                        end = q[:]
                        end[5] += delta
                        if not lower[5] <= end[5] <= upper[5]:
                            alt = q[:]
                            alt[5] -= delta
                            if lower[5] <= alt[5] <= upper[5]:
                                log(f'P{i}：J6 {delta:+d}°超限，改用反方向 {-delta:+d}°（终点位姿不变）。')
                                end, delta = alt, -delta
                            if not lower[5] <= end[5] <= upper[5]:
                                for rewound in _checked_j6_rewinds(q, lower, upper, max_deviation):
                                    if lower[5] <= rewound[5] + delta <= upper[5]:
                                        rewinds.append(rewound[:])
                                        q = rewound
                                        end = q[:]
                                        end[5] += delta
                                        break
                                else:
                                    raise ValueError(f'P{i}：J6 {delta:+d}°超限：反方向与整圈回绕均不可行。')
                        if not _fk_matches(end):
                            raise ValueError(f'P{i}：仅旋转J6无法到达所标注TCP，请检查特异点标记/工具。')
                        # v14d：换向步碰撞时，先试反方向（终点位姿不变），再试整圈回绕——
                        # TCP仿真靠方向枚举能避开这类碰撞，P2P 此前只在超限时才换向。
                        # v14j：反方向终点=当前解−delta（旧代码误算 q−2δ，朝向未翻转、FK 必不匹配，
                        # 15/15 种子全死于此——probe_p14_lookahead.py 坐实）。
                        if _movej_test_cached(q, end, 1) != 0:
                            alt = q[:]
                            alt[5] -= delta
                            flipped = False
                            if lower[5] <= alt[5] <= upper[5] and _fk_matches(alt) and _movej_test_cached(q, alt, 1) == 0:
                                log(f'P{i}：J6 {delta:+d}°扫过障碍，改用反方向 {-delta:+d}°（终点位姿不变）。')
                                end, delta, flipped = alt, -delta, True
                            if not flipped:
                                for rewound in _checked_j6_rewinds(q, lower, upper, max_deviation):
                                    cand = rewound[:]
                                    cand[5] += delta
                                    if lower[5] <= cand[5] <= upper[5] and _fk_matches(cand) and _movej_test_cached(q, cand, 1) == 0:
                                        log(f'P{i}：J6 {delta:+d}°两方向均碰，先整圈回绕再换向。')
                                        rewinds.append(rewound[:])
                                        q, end, flipped = rewound, cand, True
                                        break
                            if not flipped:
                                # v14f：两方向都碰——先切到同位姿的其他 IK 分支（碰撞预检过），
                                # 从那里再换向；途经的构型跳记入 rewinds 由执行层逐跳执行。
                                # v14j：枚举基准改为当前（未翻转）位姿——旧代码误用翻转后 target，
                                # 候选再 ±180 回到未翻转位姿，FK 对 target 永不匹配，结构性必死。
                                for cand in sorted(_ik_branch_candidates(_trajectory_pose(q), q),
                                                   key=lambda c: sum((c[j]-q[j])**2 for j in range(6))):
                                    for sgn in (delta, -delta):
                                        after = cand[:]
                                        after[5] += sgn
                                        if not (lower[5] <= after[5] <= upper[5] and _fk_matches(after)):
                                            continue
                                        if _movej_test_cached(q, cand, 1) == 0 and _movej_test_cached(cand, after, 1) == 0:
                                            log(f'P{i}：J6 ±180°两方向均碰，先切IK分支再换向（rewinds 跳转）。')
                                            rewinds.append(cand[:])
                                            q, end, delta, flipped = cand, after, sgn, True
                                            break
                                    if flipped:
                                        break
                            if not flipped:
                                # v14g：同位姿先 MoveL 到场再换向——MoveL 连续选解给出的构型
                                # 正是 TCP仿真 实测可换向的构型（贪心最近解构型两方向都扫障碍）。
                                lin_end, lin_detail = _linear_path_endpoint(q, target)
                                if lin_end is not None:
                                    pre_waypoints = _linear_waypoints(q, target)
                                    if pre_waypoints:
                                        for sgn in (delta, -delta):
                                            after = lin_end[:]
                                            after[5] += sgn
                                            if not (lower[5] <= after[5] <= upper[5] and _fk_matches(after)):
                                                continue
                                            if _movej_test_cached(lin_end, after, 1) == 0:
                                                log(f'P{i}：J6 两方向均碰，先 MoveL 到场（连续选解构型）再{sgn:+d}°换向。')
                                                plan.append(dict(method='MoveL', joints=lin_end[:], special=False,
                                                                 fallback=False, rewinds=[], j6_delta=None,
                                                                 waypoints=pre_waypoints, p2p_note='换向前MoveL到场'))
                                                q, end, delta, flipped = lin_end[:], after, sgn, True
                                                break
                            if not flipped:
                                raise ValueError(f'P{i}：J6 ±180°换向两方向均碰撞（含回绕/分支/MoveL到场尝试），该构型不可行。')
                        note = ('J6自转%+d°' % delta) if rec.get('spin360', False) else ('J6换向%+d°' % delta)
                    else:
                        target = fanuc_values_to_pose(*rec['values'])
                        # v14h：与前一点同位姿（停顿点，如轨迹7 P7）——不重新选解，
                        # 保持当前构型不动，只往计划里记一个停顿点。
                        if max(abs(_trajectory_pose(q).Pos()[j] - target.Pos()[j]) for j in range(3)) < 1e-3 and \
                           pose_angle(invH(target) * _trajectory_pose(q)) < math.radians(.01):
                            plan.append(dict(method='MoveJ', joints=q[:], special=False, fallback=False,
                                             rewinds=[], j6_delta=None, waypoints=[], p2p_note='同位姿停顿'))
                            continue
                        if not seed_used:
                            end = seed[:]  # v14c：首个TCP点直接采用种子分支（离起点可达性已在种子筛选时验证）
                            seed_used = True
                        else:
                            # v14i：前视——下一个执行点是 ±180 换向时，本点选解必须能完成那次换向
                            #（两方向任一可通行），否则贪心构型会把换向逼成死路。
                            nxt = records[i] if i < len(records) else None
                            lookahead_ok = None
                            if nxt is not None and nxt.get('singular', False) and not nxt.get('spin360', False):
                                nxt_values = nxt['values']
                                def lookahead_ok(cand, _vals=nxt_values, _lower=lower, _upper=upper):
                                    nxt_target = fanuc_values_to_pose(*_vals)
                                    for sgn in (180, -180):
                                        after = cand[:]
                                        after[5] += sgn
                                        if not (_lower[5] <= after[5] <= _upper[5]):
                                            continue
                                        err = invH(nxt_target) * _trajectory_pose(after)
                                        if norm(err.Pos()) > 1e-3 or pose_angle(err) > math.radians(.01):
                                            continue
                                        if _movej_test_cached(cand, after, 1) == 0:
                                            return True
                                    return False
                                log(f'P{i}：前视模式（P{i+1}为±180换向，选解需兼顾换向可行性）。')
                            end = (_nearest_ik_from_current_lookahead(q, target, lookahead_ok)
                                   if lookahead_ok else _nearest_ik_from_current(q, target))
                        note = 'TCP最近解直达'
                        forced_lin = False
                        # v14w24：短直线工作段强制 MoveL——P2→P3 这类 ≤210mm/姿态恒定 的
                        # 贴面平移，工艺不允许 MoveJ 关节弧绕行，直走直线（判据与直发门禁同款）。
                        # 前视夜（下一点±180换向）：直线末端同样具备换向资格才强制，否则回落
                        # MoveJ 前视绑定（保住换向可行性纪律）。
                        _rel = _trajectory_pose(q) * invH(target)
                        _seg_mm_f = norm(_rel.Pos())
                        _force_ok = _seg_mm_f <= MOVL_DIRECT_MAX_MM and pose_angle(_rel) <= math.radians(0.5)
                        # v14w33c：回撤段（TCP y 朝基座 >10mm）且下一点是同位姿换姿 ⇒ 让位 MoveJ
                        # 分支前视（强制 MoveL 的端点分支由直线 IK 连续性锁死，会对下一点无路：
                        # P5→P6→P7 实录 P7 被迫 49 跳细分）。工艺贴面滑移（Δy≈0）不受影响。
                        if _force_ok and i >= 2 and _reorient_next_pose(records, i, rec) is not None:
                            try:
                                _y_prev = float(records[i - 2]['values'][1])
                                if float(rec['values'][1]) - _y_prev > 10.0:
                                    _force_ok = False
                                    log(f'P{i}：回撤段且下一点为同位姿换姿——短直线让位 MoveJ 分支前视（v14w33c）。')
                            except Exception:
                                pass
                        if _force_ok:
                            lin_end_f, lin_detail_f = _linear_path_endpoint(q, target)
                            _lin_ok_f = (lin_end_f is not None
                                         and not _real_interfere_combo(lin_end_f)   # v14w26 组合禁区
                                         and (lookahead_ok is None or lookahead_ok(lin_end_f)))
                            if _lin_ok_f:
                                waypoints = _linear_waypoints(q, target)
                                if waypoints:
                                    end, method, fallback = lin_end_f, 'MoveL', True
                                    note = '短直线强制MoveL'
                                    forced_lin = True
                                    log(f'P{i}：短直线段（{_seg_mm_f:.1f}mm/姿态恒定）按工艺直走 MoveL（不尝试 MoveJ 弧）。')
                            elif lin_end_f is not None:
                                log(f'P{i}：短直线段直线末端无前视换向资格，回落 MoveJ 前视绑定。')
                            else:
                                log(f'P{i}：短直线段 MoveL 不可通行（{lin_detail_f}），回落 MoveJ 尝试。')
                        bound_applied = False
                        # v14j：前视绑定执行——本点是换向前夜：前视选出的构型若弧碰，不得退 MoveL
                        # （连续选解会静默锁回当前族，把死局推迟到换向步才爆——种子13 实证），
                        # 也不得由 v14c 救援收无前视资格的分支；只能换用其他前视合格分支直达，
                        # 全部失败则本构型判死、整段换种子重试。
                        if not forced_lin and lookahead_ok is not None and _movej_test_cached(q, end, 1) != 0:
                            detail_bound = _collision_details()
                            bound = None
                            for cand in sorted(_ik_branch_candidates(target, q),
                                               key=lambda c: sum((c[j]-q[j])**2 for j in range(6))):
                                if lookahead_ok(cand) and _movej_test_cached(q, cand, 1) == 0:
                                    bound = cand
                                    break
                            if bound is not None:
                                end, note, bound_applied = bound[:], '前视绑定避障直达', True
                                log(f'P{i}：前视构型弧碰（{detail_bound}），改用另一前视合格分支直达（前视绑定）。')
                            else:
                                raise ValueError(f'P{i}：MoveJ弧碰撞（{detail_bound}），其余前视合格分支均不可通行；'
                                                 '拒绝退 MoveL（连续选解会丢前视资格），本构型判死。')
                        # v14b：MoveJ 直达弧碰撞时，退回 v13 验证过的 MoveL 直线细分执行。
                        # v14w24：强制 MoveL 段不再尝试/回退 MoveJ（工艺直线优先）。
                        if not forced_lin and not bound_applied and _movej_test_cached(q, end, 1) != 0:
                            detail = _collision_details()
                            lin_end, lin_detail = _linear_path_endpoint(q, target)
                            if lin_end is None:
                                # v14c：直线也碰——枚举该目标全部 IK 分支找可通行 MoveJ（换构型救援）
                                # v14w33b：若下一点是【同位姿纯换姿】，优先选「下一点也能单条 MoveJ 贯通」
                                # 的救援分支（P6→P7 教训：P6 为自避碰选的分支对 P7 无路 ⇒ 49 跳细分拖死执行）。
                                _cands = sorted(_ik_branch_candidates(target, q),
                                                key=lambda c: sum((c[j] - q[j]) ** 2 for j in range(6)))
                                _nxt_pose = None
                                try:
                                    if i < len(records):
                                        _nr = records[i]
                                        if _nr['type'] == 'TCP' and not _nr.get('singular', False):
                                            _va = [float(v) for v in rec['values'][:6]]
                                            _vb = [float(v) for v in _nr['values'][:6]]
                                            if (all(abs(_va[k] - _vb[k]) < 1e-9 for k in range(3))
                                                    and any(abs(_va[k] - _vb[k]) > 1e-9 for k in range(3, 6))):
                                                _nxt_pose = fanuc_values_to_pose(*_nr['values'][:6])
                                except Exception:
                                    _nxt_pose = None
                                rescued = None
                                if _nxt_pose is not None:
                                    for cand in _cands:
                                        if _movej_test_cached(q, cand, 1) != 0:
                                            continue
                                        _ok_nxt = False
                                        for nb in _ik_branch_candidates(_nxt_pose, cand):
                                            if (_real_limit_ok(nb, lower, upper)
                                                    and not _real_interfere_combo(nb)
                                                    and _movej_test_cached(cand, nb, 1) == 0):
                                                _ok_nxt = True
                                                break
                                        if _ok_nxt:
                                            rescued = cand
                                            log(f'P{i}：下一点为同位姿换姿——救援分支带前视，选可与下一点单条 MoveJ 贯通的分支。')
                                            break
                                if rescued is None:
                                    for cand in _cands:
                                        if _movej_test_cached(q, cand, 1) == 0:
                                            rescued = cand
                                            break
                                if rescued is None:
                                    raise ValueError(f'P{i}：MoveJ弧碰撞（{detail}），且MoveL直线也失败：{lin_detail}；'
                                                     '该目标全部IK分支均不可通行。')
                                end, note = rescued[:], 'IK分支救援直达'
                                log(f'P{i}：最近解与直线均碰，切换IK分支救援成功。')
                            else:
                                # v14w33：同位姿/近零长（≤1mm）纯换姿段——MoveL 细分会把 90° 姿态差
                                # 切成数十跳小 MoveJ（10-21 P6→P7 实录 49 跳×每跳断连周期≈3s，
                                # 拖死执行）。优先搜无碰 MoveJ 分支单条直达（分支连续性绑死时
                                # 最近解弧碰≠无解）；搜不到再落回 MoveL 细分兜底。
                                # v14w34：_seg_mm_ro 必须是真实位置差——相对位姿平移模长在原地换姿
                                # 时被旋转杠杆放大（p−R·p，(0,-650,380) 处 90° 即 1064.8mm），
                                # 旧算式使 ≤1mm 门槛从未成立、两个搜索入口从未触发。
                                _pa = _trajectory_pose(q).Pos()
                                _pb = target.Pos()
                                _seg_mm_ro = math.sqrt(sum((_pa[_k] - _pb[_k]) ** 2 for _k in range(3)))
                                reorient_direct = None
                                if _seg_mm_ro <= 1.0:
                                    for cand in sorted(_ik_branch_candidates(target, q),
                                                       key=lambda c: sum((c[j]-q[j])**2 for j in range(6))):
                                        if (not _real_interfere_combo(cand)
                                                and _real_limit_ok(cand, lower, upper)
                                                and (lookahead_ok is None or lookahead_ok(cand))
                                                and _movej_test_cached(q, cand, 1) == 0):
                                            reorient_direct = cand
                                            break
                                if reorient_direct is not None:
                                    end, note = reorient_direct[:], '同位姿换姿MoveJ直达'
                                    method, fallback = 'MoveJ', False
                                    waypoints = []
                                    log(f'P{i}：同位姿换姿——MoveL 细分会碎成数十小段，改用无碰 MoveJ 分支单条直达。')
                                elif _seg_mm_ro <= 1.0 and plan and rec['type'] == 'TCP' and i >= 2:
                                    # v14w33d：回改上一步（已入计划、未执行）为可与本点单条 MoveJ 贯通的
                                    # 分支——上一步若走最近解直达/救援，其分支未必对本点有路（P6→P7 实录）。
                                    # 改关节目标后两跳路径均当场重检，证书完整。
                                    _prev_step = plan[-1]
                                    _prev_q = _prev_step['joints']
                                    _prev_prev = plan[-2]['joints'] if len(plan) >= 2 else saved
                                    _prev_pose = fanuc_values_to_pose(*records[i - 2]['values'][:6])
                                    reorient_direct = None
                                    for c6 in sorted(_ik_branch_candidates(_prev_pose, _prev_prev),
                                                     key=lambda c: sum((c[k] - _prev_q[k]) ** 2 for k in range(6))):
                                        if _real_interfere_combo(c6) or not _real_limit_ok(c6, lower, upper):
                                            continue
                                        if _movej_test_cached(_prev_prev, c6, 1) != 0:
                                            continue
                                        for c7 in sorted(_ik_branch_candidates(target, c6),
                                                         key=lambda c: sum((c[k] - c6[k]) ** 2 for k in range(6))):
                                            if _real_interfere_combo(c7) or not _real_limit_ok(c7, lower, upper):
                                                continue
                                            if lookahead_ok is not None and not lookahead_ok(c7):
                                                continue
                                            if _movej_test_cached(c6, c7, 1) != 0:
                                                continue
                                            _prev_step['joints'] = c6[:]
                                            reorient_direct = c7
                                            break
                                        if reorient_direct is not None:
                                            break
                                    if reorient_direct is not None:
                                        end, note = reorient_direct[:], '同位姿换姿MoveJ直达'
                                        method, fallback = 'MoveJ', False
                                        waypoints = []
                                        log(f'P{i}：回改上一步分支后，本点取得单条 MoveJ 直达（两跳均重检无碰）。')
                                if reorient_direct is not None:
                                    pass   # 已在上方处理
                                else:
                                    waypoints = _linear_waypoints(q, target)
                                    if not waypoints:
                                        raise ValueError(f'P{i}：MoveJ弧碰撞（{detail}），MoveL细分采样失败，拒绝。')
                                    end, method, fallback = lin_end, 'MoveL', True
                                    note = 'MoveJ弧碰退回MoveL细分'
                                    log(f'P{i}：MoveJ弧碰撞（{detail}），改走 MoveL 直线细分（{len(waypoints)} 途经点）。')
                    if not all(lower[j] <= end[j] <= upper[j] for j in range(6)):
                        raise ValueError(f'P{i}：关节超限，J6目标={end[5]:.3f}°。')
                    if method == 'MoveJ' and _movej_test_cached(q, end, 1) != 0:
                        # v14e：普通TCP点最后一级救援——v13 遗产 _obstacle_joint_target
                        # （21候选、肘高排序、限TCP偏离）选避障构型，TCP仿真靠它在同一站过关。
                        try:
                            end = _obstacle_joint_target(q, rec['values'], max_deviation, log)
                            note = '避障选解直达'
                        except ValueError:
                            raise ValueError(f'P{i}：MoveJ路径检查失败（含避障选解）：' + _collision_details())
                        if _movej_test_cached(q, end, 1) != 0:
                            raise ValueError(f'P{i}：MoveJ路径检查失败：' + _collision_details())
                    # v14w25：J6 恰=±360 边界值被控制器 -40006 拒收（10-15 17:26/17:33 实录）。
                    # v14w32：±359.999 内推仍防不住「J6 单轴被丢弃」（10-21 P4 实证：J1~J5 全到、
                    # J6 纹丝停在 180、误差 180°）——改为换 (−180,180] 同角表示（359.999→−0.001），
                    # J6 彻底离开 ±360 邻域。换表示会翻转 MoveJ 弧方向 ⇒ 必须重检路径，不过即报规划错误。
                    # spin360/多圈值（|J6|>360.001）不在此列，防绞坏自转语义。
                    if abs(end[5]) >= 359.999 and abs(end[5]) <= 360.001 and not rec.get('spin360'):
                        _j6n = end[5] - math.copysign(360.0, end[5])
                        log(f'P{i}：J6={end[5]:.3f}° 贴 ±360 边界，换同角表示 {_j6n:.3f}°（v14w32：±359.999 仍被丢轴，彻底离开边界邻域）。')
                        end[5] = _j6n
                        for _wp in waypoints:
                            if abs(_wp[5]) >= 359.999 and abs(_wp[5]) <= 360.001:
                                _wp[5] = _wp[5] - math.copysign(360.0, _wp[5])
                        if method == 'MoveJ' and _movej_test_cached(q, end, 1) != 0:
                            raise ValueError(f'P{i}：J6 换同角表示后 MoveJ 路径碰撞：' + _collision_details())
                    # v14w26：解落入实机自干涉组合区（J4×J5，-40006）——MoveJ 解自动换无碰安全
                    # 分支直达；直线段落区（强制/兜底）整段换种子；无安全分支则判死。
                    if _real_interfere_combo(end):
                        if method == 'MoveJ' and rec['type'] == 'TCP' and not rec.get('singular', False):
                            rescued_if = None
                            for cand_if in sorted(_ik_branch_candidates(target, q),
                                                   key=lambda c: sum((c[j]-q[j])**2 for j in range(6))):
                                if (_real_limit_ok(cand_if, lower, upper)
                                        and not _real_interfere_combo(cand_if)
                                        and _movej_test_cached(q, cand_if, 1) == 0):
                                    rescued_if = cand_if
                                    break
                            if rescued_if is None:
                                raise ValueError(f'P{i}：全部无碰分支均落入实机自干涉组合区'
                                                 f'（|J4|>{REAL_INTERFERE_J4_MAX:.0f} 且 |J5|>{REAL_INTERFERE_J5_MIN:.0f}，-40006 实录区），本构型判死。')
                            log(f'P{i}：预选解落入实机自干涉组合区（J4={end[3]:.1f}°, J5={end[4]:.1f}°），换安全分支直达。')
                            end = rescued_if[:]
                            note = '自干涉安全分支直达'
                        else:
                            raise ValueError(f'P{i}：该步解落入实机自干涉组合区（J4={end[3]:.1f}°, J5={end[4]:.1f}°），换种子重试。')
                    plan.append(dict(method=method, joints=end[:], special=rec.get('singular', False), fallback=False,
                                     rewinds=rewinds, j6_delta=delta,
                                     waypoints=waypoints, p2p_note=note))
                    q = end[:]
                if _continuous_profile_active:
                    previous = saved
                    for number, step in enumerate(plan, 1):
                        if step.get('waypoints'):
                            rel = _trajectory_pose(step['joints']) * invH(_trajectory_pose(previous))
                            if (step['method'] != 'MoveL' or norm(rel.Pos()) > MOVL_DIRECT_MAX_MM
                                    or pose_angle(rel) > math.radians(.5)):
                                raise ValueError(f'P{number}将退回{len(step["waypoints"])}段停走，换入口分支重试。')
                        previous = step['joints']
                log('逐段规划完成，开始整段碰撞复核（1mm/1°采样，请稍候）…')
                _verify_obstacle_plan(saved, plan)
                _certify_continuous_direct(records, saved, plan, log)
                _preferred_seed = (seed_context, seed)
                log(f'P2P+奇异点整段路径预检通过：{len(plan)}点。')
                return plan
            except ValueError as exc:
                last_seed_error = exc
                log(f'种子 {seed_rank}/{len(seeds)} 在此构型失败（{exc}），换下一构型整段重试…')
        if last_seed_error is not None:
            raise last_seed_error
    finally:
        _continuous_profile_active = False
        robot.setJoints(saved)
        RDK.Render(True)

root = tk.Tk()
root.title("RoboDK - 机械臂运动控制（P2P v15.21）")
root.geometry("1200x750")
root.resizable(True, True)

tk.Label(root, text="Dobot CR5 运动控制", font=("Microsoft YaHei", 16, "bold")).pack(pady=10)

notebook = ttk.Notebook(root)
notebook.pack(fill=tk.BOTH, expand=True, padx=10, pady=5)

# ---- 选项卡 1：单点运动 ----
tab_single = ttk.Frame(notebook)
notebook.add(tab_single, text="单点运动")

frame_coord = tk.LabelFrame(tab_single, text="目标 TCP（Fanuc 格式）")
frame_coord.pack(fill=tk.X, padx=10, pady=10)

names = ["X (mm)", "Y (mm)", "Z (mm)", "Rx (deg)", "Ry (deg)", "Rz (deg)"]
defaults = ["0.000", "-241.500", "1047.000", "-90.000", "0.000", "180.000"]
entries_single = []

for i in range(6):
    tk.Label(frame_coord, text=names[i]).grid(row=0, column=i*2, padx=5, pady=10)
    e = tk.Entry(frame_coord, width=12)
    e.insert(0, defaults[i])
    e.grid(row=0, column=i*2+1, padx=5, pady=10)
    entries_single.append(e)

frame_mtype = tk.Frame(tab_single)
frame_mtype.pack(fill=tk.X, padx=10, pady=5)
move_type = tk.StringVar(value="MoveL")
tk.Radiobutton(frame_mtype, text="MoveL (直线)", variable=move_type, value="MoveL").pack(side=tk.LEFT, padx=10)
tk.Radiobutton(frame_mtype, text="MoveJ (关节)", variable=move_type, value="MoveJ").pack(side=tk.LEFT, padx=10)

btn_single_frame = tk.Frame(tab_single)
btn_single_frame.pack(fill=tk.X, padx=10, pady=5)

def _read_current():
    read_current(entries_single)
def _fill_current():
    fill_current(entries_single)
def _check_ik():
    check_ik_single(entries_single)
def _exec_single():
    execute_single(entries_single, move_type.get())

tk.Button(btn_single_frame, text="读取当前 TCP", command=_read_current, width=15).pack(side=tk.LEFT, padx=3)
tk.Button(btn_single_frame, text="当前 TCP -> 输入框", command=_fill_current, width=20).pack(side=tk.LEFT, padx=3)
tk.Button(btn_single_frame, text="检测可达性", command=_check_ik, width=15, bg="#2196F3", fg="white").pack(side=tk.LEFT, padx=3)
tk.Button(btn_single_frame, text="执行运动", command=_exec_single, width=20,
          font=("Microsoft YaHei", 10, "bold"), bg="#4CAF50", fg="white").pack(side=tk.LEFT, padx=3)


# ---- 选项卡 2：目标关节运动（实机） ----
tab_joint = ttk.Frame(notebook)
notebook.add(tab_joint, text="目标关节运动")

frame_joint = tk.LabelFrame(tab_joint, text="目标关节（deg）")
frame_joint.pack(fill=tk.X, padx=10, pady=10)

joint_names = ["J1 (deg)", "J2 (deg)", "J3 (deg)", "J4 (deg)", "J5 (deg)", "J6 (deg)"]
joint_defaults = ["0.000", "0.000", "0.000", "0.000", "0.000", "0.000"]
entries_joint = []

for i in range(6):
    tk.Label(frame_joint, text=joint_names[i]).grid(row=0, column=i*2, padx=5, pady=10)
    e = tk.Entry(frame_joint, width=12)
    e.insert(0, joint_defaults[i])
    e.grid(row=0, column=i*2+1, padx=5, pady=10)
    entries_joint.append(e)

btn_joint_frame = tk.Frame(tab_joint)
btn_joint_frame.pack(fill=tk.X, padx=10, pady=8)

def _read_current_joint_values():
    read_current_joints(entries_joint)

def _fill_current_joints():
    fill_current_joints(entries_joint)

def _exec_joint():
    execute_joint_target(entries_joint)

def _zero_joints():
    clear_joint_target(entries_joint)

tk.Button(btn_joint_frame, text="读取当前关节", command=_read_current_joint_values, width=14).pack(side=tk.LEFT, padx=3)
tk.Button(btn_joint_frame, text="当前关节 -> 输入框", command=_fill_current_joints, width=20).pack(side=tk.LEFT, padx=3)
tk.Button(btn_joint_frame, text="执行指定关节 MoveJ", command=_exec_joint, width=24,
          font=("Microsoft YaHei", 10, "bold"), bg="#FF9800", fg="white").pack(side=tk.LEFT, padx=3)
tk.Button(btn_joint_frame, text="清零", command=_zero_joints, width=10).pack(side=tk.LEFT, padx=3)

tk.Label(tab_joint,
         text="输入 J1~J6 目标角度（deg）；完整关节路径预检通过后才发送实机 MoveJ。",
         fg="#555555").pack(anchor=tk.W, padx=15, pady=5)
tk.Label(tab_joint,
         text="安全提示：首次测试建议只改变一个关节、改变 5~10°，确认方向和角度定义正确后再进行大角度运动。",
         fg="#C62828").pack(anchor=tk.W, padx=15, pady=2)

# ---- 选项卡 3：连续运动 ----
tab_traj = ttk.Frame(notebook)
notebook.add(tab_traj, text="连续运动")

frame_traj_input = tk.LabelFrame(
    tab_traj,
    text="连续运动点输入：每次输入 1 个 TCP 点或 1 组关节角度，点击“检查并加入”"
)
frame_traj_input.pack(fill=tk.X, padx=10, pady=10)

type_frame = tk.Frame(frame_traj_input)
type_frame.pack(fill=tk.X, padx=8, pady=5)

tk.Label(type_frame, text="点类型：").pack(side=tk.LEFT, padx=3)

traj_type = tk.StringVar(value="TCP")
tk.Radiobutton(
    type_frame, text="TCP（X,Y,Z,Rx,Ry,Rz）",
    variable=traj_type, value="TCP"
).pack(side=tk.LEFT, padx=8)

tk.Radiobutton(
    type_frame, text="关节（J1~J6）",
    variable=traj_type, value="JOINT"
).pack(side=tk.LEFT, padx=8)

traj_names_tcp = ["X", "Y", "Z", "Rx", "Ry", "Rz"]
traj_names_joint = ["J1", "J2", "J3", "J4", "J5", "J6"]

traj_entries = []

# ---- 末端特异点设置 ----
singular_var = tk.BooleanVar(value=False)
j6_direction_var = tk.IntVar(value=180)

singular_frame = tk.Frame(frame_traj_input)
singular_frame.pack(fill=tk.X, padx=8, pady=3)

tk.Checkbutton(
    singular_frame,
    text="末端特异点（跳过IK，仅J6转动）",
    variable=singular_var
).pack(side=tk.LEFT, padx=3)

tk.Label(singular_frame, text="J6方向：").pack(side=tk.LEFT, padx=(15, 3))
tk.Radiobutton(singular_frame, text="+180°", variable=j6_direction_var, value=180).pack(side=tk.LEFT, padx=3)
tk.Radiobutton(singular_frame, text="-180°", variable=j6_direction_var, value=-180).pack(side=tk.LEFT, padx=3)
spin_var = tk.BooleanVar(value=False)
tk.Checkbutton(singular_frame, text="J6自转360°（第二类，六维与前点相同）", variable=spin_var).pack(side=tk.LEFT, padx=3)

# 输入框单独放在 grid 子容器中。
# frame_traj_input 本身使用 pack 管理子控件，不能再直接对它的子控件使用 grid。
traj_value_frame = tk.Frame(frame_traj_input)
traj_value_frame.pack(fill=tk.X, padx=8, pady=5)

for i in range(6):
    tk.Label(
        traj_value_frame,
        text=traj_names_tcp[i]
    ).grid(row=0, column=i * 2, padx=3, pady=8)

    e = tk.Entry(traj_value_frame, width=12)
    e.grid(row=0, column=i * 2 + 1, padx=4, pady=8)
    traj_entries.append(e)

# 默认先按 TCP 输入显示
tcp_defaults = ["0.000", "-241.500", "1047.000", "-90.000", "0.000", "180.000"]
for e, val in zip(traj_entries, tcp_defaults):
    e.insert(0, val)


def _update_traj_labels_and_defaults():
    """切换 TCP/关节输入时，更新标签和默认值。"""
    names = traj_names_tcp if traj_type.get() == "TCP" else traj_names_joint
    defaults = (
        tcp_defaults
        if traj_type.get() == "TCP"
        else ["0.000"] * 6
    )

    for i, e in enumerate(traj_entries):
        # grid 上的 Label 位于当前列
        for widget in traj_value_frame.grid_slaves(row=0, column=i * 2):
            widget.configure(text=names[i])

        e.delete(0, tk.END)
        e.insert(0, defaults[i])


tk.Radiobutton(
    type_frame, text="TCP（X,Y,Z,Rx,Ry,Rz）",
    variable=traj_type, value="TCP",
    command=_update_traj_labels_and_defaults
).pack_forget()

# 重新建立带 command 的两个单选按钮
for widget in list(type_frame.pack_slaves()):
    if isinstance(widget, tk.Radiobutton):
        widget.destroy()

tk.Radiobutton(
    type_frame, text="TCP（X,Y,Z,Rx,Ry,Rz）",
    variable=traj_type, value="TCP",
    command=_update_traj_labels_and_defaults
).pack(side=tk.LEFT, padx=8)

tk.Radiobutton(
    type_frame, text="关节（J1~J6）",
    variable=traj_type, value="JOINT",
    command=_update_traj_labels_and_defaults
).pack(side=tk.LEFT, padx=8)

btn_traj_input = tk.Frame(tab_traj)
btn_traj_input.pack(fill=tk.X, padx=10, pady=3)

tk.Button(
    btn_traj_input,
    text="检查并加入当前点",
    command=add_and_check_trajectory_point,
    width=22,
    bg="#2196F3",
    fg="white",
    font=("Microsoft YaHei", 10, "bold")
).pack(side=tk.LEFT, padx=3)

tk.Button(
    btn_traj_input,
    text="读取当前TCP并写入",
    command=read_current_tcp_to_traj,
    width=20
).pack(side=tk.LEFT, padx=3)

tk.Button(
    btn_traj_input,
    text="读取当前关节并写入",
    command=read_current_joints_to_traj,
    width=20
).pack(side=tk.LEFT, padx=3)

tk.Button(
    btn_traj_input,
    text="清空当前输入",
    command=clear_trajectory_input,
    width=16
).pack(side=tk.LEFT, padx=3)

tk.Label(
    tab_traj,
    text="加入点时检查格式并保留关节圈数；执行前再进行整段限位、台子和地面碰撞检查。",
    fg="#555555"
).pack(anchor=tk.W, padx=15, pady=3)

frame_record = tk.LabelFrame(
    tab_traj,
    text="已检查通过的连续运动点（按加入顺序执行，可混合 TCP / 关节点）"
)
frame_record.pack(fill=tk.BOTH, expand=True, padx=10, pady=8)

record_text = tk.Text(frame_record, font=("Consolas", 10), height=10)
record_text.pack(fill=tk.BOTH, expand=True, padx=5, pady=5)

btn_record_frame = tk.Frame(tab_traj)
btn_record_frame.pack(fill=tk.X, padx=10, pady=4)

tk.Button(
    btn_record_frame, text="删除最后一点",
    command=delete_last_record, width=15
).pack(side=tk.LEFT, padx=3)

tk.Button(
    btn_record_frame, text="清空全部点",
    command=clear_records, width=15
).pack(side=tk.LEFT, padx=3)

tk.Button(
    btn_record_frame, text="导入轨迹",
    command=import_trajectory, width=14
).pack(side=tk.LEFT, padx=3)

tk.Button(
    btn_record_frame, text="执行整段连续运动",
    command=execute_recorded_trajectory,
    width=24,
    font=("Microsoft YaHei", 10, "bold"),
    bg="#4CAF50", fg="white"
).pack(side=tk.LEFT, padx=3)

tk.Label(
    tab_traj,
    text="执行前按实机当前关节完成台子/地面预检；仅执行已验证方案。驱动报断连时复核实际到位；未到位或其他异常时中止。",
    fg="#555555"
).pack(anchor=tk.W, padx=15, pady=4)

real_deviation_var = tk.StringVar(value="500.0")
frame_deviation = tk.Frame(root)
frame_deviation.pack(fill=tk.X, padx=10, pady=3)
tk.Label(frame_deviation, text="预检MoveJ兜底最大TCP偏离(mm)：").pack(side=tk.LEFT)
tk.Entry(frame_deviation, textvariable=real_deviation_var, width=10).pack(side=tk.LEFT)
tk.Label(frame_deviation, text="默认500：与TCP仿真/轨迹7~11验证口径一致；实机速度10 mm/s（v14w25 调慢）").pack(side=tk.LEFT, padx=8)

# v14w24：法兰补偿MOVL 默认开启，勾选框移除（工艺定型）。v14l 实机判决驱动 MOVL 无工具
# 补偿（按法兰执行，无补偿直发已拉黑勿回归）；v14p 将错就错把法兰位姿当笛卡尔目标直发，
# 法兰被精确送达→物理尖端走在认证直线上。v14w36/37：位姿由调用方自算 invH(PoseFrame)*SolveFK
# （动画=认证直线，根治关节弧假碰撞冻死），发送窗口配单位变换（校验/数字=法兰空间）。
# 适用：MoveL 细分段≤210mm 且姿态恒定（v14w35 门禁）；规划/预检/几何零改动；失败指纹照旧即停；净化失败自动回落细分。
real_movldirect_var = tk.BooleanVar(value=True)   # 仅保留变量接口（执行入口读取）；无 GUI 控件

# ---- 日志区 ----
frame_log = tk.LabelFrame(root, text="日志")
frame_log.pack(fill=tk.BOTH, expand=True, padx=10, pady=5)

text_log = scrolledtext.ScrolledText(frame_log, font=("Consolas", 10), height=8)
text_log.pack(fill=tk.BOTH, expand=True, padx=5, pady=5)

# ============================================================
# 启动
# ============================================================
log("机器人: " + robot.Name())
log("程序就绪。" + LOG_VERSION + " ｜ 模式：RUNMODE_RUN_ROBOT + robot.Connect() ｜ 文件日志：" + LOG_PATH)
_ensure_canonical_tool()   # v14w17：启动守护（覆盖"加载了带归零工具的存档"场景）
log("单点：输入坐标 -> 检测可达性 -> 执行 MoveL/MoveJ")
log("目标关节：输入 J1~J6 -> 实机 MoveJ（不经过 TCP/Fanuc 转换和 IK）")
log("连续运动（P2P v15.21）：修改点位后仍启用分支搜索、防停走及逐段重新认证；无法认证的直线在发送运动前停止；130mm TCP。")

def _log_pump():
    try:
        while True:
            text_log.insert(tk.END, _log_queue.get_nowait() + NL)
            text_log.see(tk.END)
    except Exception:
        pass
    root.after(100, _log_pump)


_close_requested = False


def _idle_tool_guard():
    if not _real_running and not _tool_window_depth:
        try:
            if _same_tool_pose(robot.PoseTool(), eye(4)):
                _ensure_canonical_tool()
            if _close_requested:
                root.destroy()
                return
        except Exception as exc:
            _file_log('工具空闲守护失败：' + str(exc))
    root.after(1000, _idle_tool_guard)


def _on_close():
    global _close_requested
    if _real_running:
        _close_requested = True
        log('已请求关闭：等待当前任务结束并恢复 TCP 后关闭窗口，继续保留到位监控。')
        return
    _ensure_canonical_tool()
    root.destroy()


root.protocol('WM_DELETE_WINDOW', _on_close)
root.after(100, _log_pump)
root.after(1000, _idle_tool_guard)
_start_heartbeat()
try:
    root.mainloop()
except BaseException:
    import traceback
    _file_log('FATAL mainloop: ' + traceback.format_exc())
    raise

--- program _TCP仿真_路径预检 ---

--- Python program TCP真实运动_P2P版 ---
# -*- coding: utf-8 -*-
"""
RoboDK 实机运动控制（基于 robodk_movej_diag.py 的成功模式）
- 单点：TCP 输入 -> IK 检测 -> MoveL/MoveJ 执行
- 连续轨迹：与TCP仿真同款（姿态退让、J6特异点±180°/自转360°、避障规划+缓存）
2026-10-09：连续运动逻辑对齐 机械臂TCP仿真_副本.py；预检偏离默认 50→500（与验证口径一致）
模式：RUNMODE_RUN_ROBOT + robot.Connect()
"""

from robodk.robolink import *
from robodk.robomath import *
import tkinter as tk
from tkinter import ttk, scrolledtext, filedialog
import time
import math
import json
import itertools

ROBOT_SPEED = 10.0   # v14w25：20→10 mm/s（用户要求调慢；顺带拉长指令间隔，缓解驱动掉线-重连压力）
CANONICAL_TOOL = (0.0, 0.0, 130.0, 0.0, 0.0, 0.0)   # v14w40：规范工具 182→126（2026-10-23 最终实测 法兰→TCP=126；v14w27~39 为 182、v14w14~w26 为 100）；守护用
NL = chr(10)
import queue as _queue_mod
_log_queue = _queue_mod.Queue()  # 后台线程日志经队列回流主线程，GUI 不冻结
LOG_PATH = r'D:\mydata\glm-workplace\sim_scripts\real_gui_log_p2p.txt'  # P2P版独立日志，不覆盖v13黑匣子
LOG_VERSION = 'v15.22-20261104'   # ★ 版本号规则（用户 2026-11-03 要求）：【每次改动都要升版本号】
                               # v15   ：从 v14w42 更名（J4 150→178 / P9 入禁直发 / Tool-User 实验开关 / 删超长横幅）
                               # v15.1 ：最后防线同角归一化修复（段6 J4=198.78 ≡ −161.22 被误判超限）
                               # v15.2 ：新增 |J4|>150 单独硬禁区（治 P5 的 J4=172.88 姿态自干涉）
                               # v15.3 ：打开 MOVL_SEND_TOOL_USER（直发前发 Tool(0)/User(0)，验证能否根治断断续续）
                               # v15.4 ：收口 MoveJ 加重试（治 P8 停下：收口遇断连没走完 ⇒ 关节残差 2.68° 残留）
                               # v15.5 ：直发+收口后再做【关节校正重试】（治 P8 停下：收口走假断连分支 ⇒ 报"已完成"但关节没到位）
                               # v15.6 ：_require_joints 改【带重试的稳定判定】（治 P8 尾通过 → P9 开头又失败：中间还在微动）
                               # v15.7 ：直发后先等【关节真静止】再做验收/收口（治 P8 的 elbow-flip 假通过/假失败）
                               # v15.8 ：★直发落点【自干涉安全网】—— 控制器自行选解可能落进禁区 ⇒ 立刻回认证构型
                               # v15.9 ：P8 也禁直发（治"选解自由"：J1/J6 同步偏 9.77° = 另一组 IK 解）⇒ P8 走细分
                               # v15.10：_require_joints 失败时【主动发 MoveJ 校正】（根治 P8 后不动：断连分支对 MoveJ 只等静止不等到位）
                               # 下次改动 ⇒ v15.23；标题与下方"连续运动"横幅要同步改
# v14w41：独立命名 TCP/法兰工具；恢复原工具链接并核验，失败停止；空闲守护与延后关闭。
# 历史版本记录（场景坐标并非实时状态）：★ v14w40（2026-10-23 18:09）：工具定案 126——最终实测 法兰→TCP=126，CANONICAL_TOOL/守护恢复值/banner 同步 126（历史：v14w27~39=182、v14w14~26=100）；配套场景 磨砂圆柱 y −860→−886、挡板 y 56→30（整体 −26 抵消工具加长的 26mm 深度偏移），轨迹13 采用 z460 统一版（连续轨迹13_t126_z460.json）——tool126+z460+场景−26 组合实测预检 21/21 PASS。⚠️ 实物圆柱/挡板须同步 −26；面贴滚轮旧坐标全部失效需重解；轨迹14/15 需在新配置下复验。v14w39（2026-10-22 14:31）：flange 窗口（单位变换+藏把手）从「仅包 RPC」扩大到【覆盖整个 settle 生命周期】。v14w38 失败教训：假断连让 MoveL 调用秒抛、窗口当场关闭、把手提前恢复，而真实滑行+RoboDK 本地退化动画仍在跑——本地动画在弧 66% 被碰撞检测掐停（模型冻点 J1≈67 四次实录同一位置）、红显常驻，收口 MoveJ 从撞点姿态发出被 RoboDK 拦死。v14w39 三件套：①窗口=包装层全程（发送+断连恢复+到位等待，补发重试每次重开窗）；②守卫补恢复隐藏态门把手（防 GUI 中杀留下隐藏态污染预检）；③直发 settle 返回后 robot.setJoints 钉模型到认证终点（清残余态双保险）。真直线 1mm 检查 0 碰撞、柜子零报警不变。v14w38：窗口藏把手（范围不足判负）。v14w37：位姿传递+单位变换（P8 TargetReachError 修复）。v14w35：门禁 210。v14w34：_seg_mm_ro 真位置差。其余见前版注释与 MEMORY。
# v14w32（2026-10-21 10:58）：J6 贴 ±360 边界的处置从「±359.999 内推」改为「换 (−180,180] 同角表示」（359.999→−0.001）——10-21 P4 实证：内推值仍被控制器丢 J6 单轴（J1~J5 全到、J6 停在 180、误差 180°）；换表示后当场重检 MoveJ 路径（方向翻转风险）；spin360/|J6|>360.001 不处理。其余=v14w30（阈值5°；v14w31 已撤回）。
# v14w30（2026-10-21 09:31）：MovL 直发到位阈 MOVL_ARRIVE_TOL_DEG 2°→5°——10-21 P8 实证：tool=182+z=380 构型下控制器 ~5mm 固有落点误差映射为关节 2.58°（tool=100 时代仅 0.7~0.9°），卡死在旧 ≤2° 阈值外被误判"疑似未执行"；臂实为完成态（零速/模式5/无报警）。护栏不降级：法兰级粗验收(≤8mm/≤1°)+MoveJ 收口仍在其后罩终点；60s 上限与不重发不变。（v14w31 稳定窗+补发×3 已于 10-21 按用户要求撤回。）
# v14w29（2026-10-20 16:42）：站内 圆柱+挡板 统一后移（远离基座）82mm（用户指令：尖端距圆柱面仅 14mm 太近、易自干涉）——圆柱 pose.y −840→−922、挡板 pose.y 76→−6；同时修正 10-15 起过期的场景注释。轨迹13 六点 z−82 补丁后离线预检 21/21 全绿（含本次场景移动复验）。
# v14w28（2026-10-20 16:15）：网格注释同步（纯注释版，逻辑零改动）——把手网格手术 v4：连接件加长、把手组件整体外移，【把手工作点=法兰前 182mm】，stl=tools\handle_rod_182_v2.stl（站内已换、未保存）。工具仍=182mm。
# v14w27（2026-10-20 15:49）：工具坐标 100→182mm（用户实测【物理工具真实长度】；站内 PoseTool 已同步 [0,0,182]）——CANONICAL_TOOL/守护恢复值/直发注释同步，全部 IK 按 182 解算。⚠️ 轨迹13 有 5 点（P8/P9/P10/P12/P13）在 182 下超臂展无逆解，重新示教前禁实机。
# v14w26（2026-10-15 18:15）：实机自干涉组合区（PoseSelfInterference 的 J4×J5 耦合，-40006 实录）——J4=-115.5×J5=173.1 与 J4=-109.4×J5=171.5 双拒；安全实录 J4=-83.2×J5=177.6。修：规划期禁选 |J4|>100 且 |J5|>165 的组合（MoveJ 解落区自动换无碰安全分支；直线段落区回落；无安全分支则整段换种子）。沿用 v14w25：速度10mm/s、J6±360内推（保留作防御）；v14w24：短直线强制MoveL、直发默认开。
# v14w20：受控补发。v14w19：三角离零域。v14w17：工具守护。工具=182.000（v14w27 起）；把手网格=v4 手术（把手组件外移、工作点 z=182，尖端=TCP，把手端抓手 z∈[174,182]；v14w28 起 stl=handle_rod_182_v2）。
# 场景（2026-10-20 实测，v14w29 圆柱/挡板统一后移82 后）：圆柱（轴∥X 滚轮 R150×H50）世界包络 X[−25,25] Y[−1062,−782] Z[330,610]；挡板世界包络 X[−235,215] Y[−1232,−932] Z[150,900]。10-13 版旧场景注释坐标已废（10-15 起站内多次平移未同步注释，v14w29 起以本行为准）。
# 控制器日志实锤（logs/all/log）：
#   11:38:20 拒收 MovL(-0.000000,-615.371000,300.000000,90.000000,0.000000,-0.000000)
#            → [MovL#820] the type of params is wrong: -30001 —— 这才是 P9 直发 60s 零位移的真凶；
#   15:55:51 单步同目标接受 MovL(0.000000,-615.371000,299.999986,89.999995,-0.000003,0.000000)
#            → return 0，1.1s 到位、法兰验收 5.08mm/0.61° 过。两样本差在【边界形态】：
#            x 负零/极小负、rx 恰=+90.000000、rz 负零（触发器三候选未最终定死，净化同时设防）。
# 修法：直发前 _movl_digit_safe_joints 只在零附近边界区对发送关节微扰（单关节 ≤0.05°、末端 ≲0.6mm
#   ≪ 圆柱真裕度 19.9mm）；到位/法兰验收/MoveJ 收口仍全部对【原始认证关节】判定，收口回认证构型。
#   净化失败 ⇒ 本段自动改走细分途经点（安全回落，不比 v14u 更糟）。
# 备份：…_v14v4_20261013-1608.py.bak（另有 1208 站内导出副本）；v14v/v2/v3 回退项见 P2P_LESSONS.md。
# 旧 v14u 备注：v14t 10:38 复跑判读——P9 起步延迟 >6s，「起点静止」与「完成静止」反馈不可区分，位置对目标才是唯一可靠锚点
# v12 黑匣子：原生崩溃时把 Python 调用栈转储到独立文件（被动，不影响逻辑）
# 注意：faulthandler.enable 只接受文件对象，传路径字符串会 AttributeError（v12 首版踩坑，已被 except 吞掉）
CRASH_PATH = r'D:\mydata\glm-workplace\sim_scripts\real_gui_crash.txt'
try:
    import faulthandler as _fh
    _crash_fp = open(CRASH_PATH, 'a', encoding='utf-8')
    _fh.enable(_crash_fp, all_threads=True)
except Exception:
    pass

def _file_log(s):
    try:
        import io as _io, time as _time
        with _io.open(LOG_PATH, 'a', encoding='utf-8') as f:
            f.write(_time.strftime('%m-%d %H:%M:%S') + ' | ' + str(s) + NL)
    except Exception:
        pass


RDK = Robolink()

def fanuc_to_pose(x, y, z, rx, ry, rz):
    return Fanuc_2_Pose([x, y, z, rx, ry, rz])

def pose_to_fanuc(pose):
    return Pose_2_Fanuc(pose)

# ---- 获取机器人 ----
robot = RDK.Item('Dobot CR5', ITEM_TYPE_ROBOT)
if not robot.Valid():
    raise Exception("未找到机器人")

# ---- 全局变量 ----
text_points = None
text_log = None
record_text = None
entries_single = None
entries_joint = None
move_type = None
trajectory_records = []
_connected = False

# ============================================================
# 日志
# ============================================================
# v12 心跳：每5秒覆写一次小文件（时间戳+pid+日志末行），进程死亡时间一目了然
HEARTBEAT_PATH = r'D:\mydata\glm-workplace\sim_scripts\real_gui_heartbeat.txt'

def _start_heartbeat():
    import threading as _t, time as _time, os as _os, io as _io
    def _beat():
        while True:
            try:
                last = ''
                try:
                    with _io.open(LOG_PATH, 'r', encoding='utf-8') as f:
                        _lines = f.read().splitlines()
                        last = _lines[-1] if _lines else ''
                except Exception:
                    pass
                with _io.open(HEARTBEAT_PATH, 'w', encoding='utf-8') as f:
                    f.write('%s | pid=%d | alive\nlast: %s\n' % (
                        _time.strftime('%m-%d %H:%M:%S'), _os.getpid(), last[:150]))
            except Exception:
                pass
            _time.sleep(5.0)
    _t.Thread(target=_beat, daemon=True, name='gui_heartbeat').start()


def log(s):
    _file_log(s)  # 先落盘：即使后续 print 阻塞，磁盘日志也不受影响
    print(s)
    if text_log:
        try:
            _log_queue.put_nowait(str(s))
        except Exception:
            text_log.insert(tk.END, str(s) + NL)

# ============================================================
# 连接（只连一次，复用）
# ============================================================
def ensure_connected():
    global _connected
    try:
        status, msg = robot.ConnectedState()
        if status != ROBOTCOM_READY:
            if status >= 0:
                log('机器人未就绪，取消执行：' + str(msg))
                return False
            robot.Connect()
            # v14o：固定 1.5s 改为就绪探测（0.3s 轮询，最多 3s）：假断连恢复是每跳尾部
            # 停顿税的一部分；探测到就绪即返回，未就绪语义与旧版一致（返回 False）。
            for _ in range(10):
                time.sleep(0.3)
                status, msg = robot.ConnectedState()
                if status == ROBOTCOM_READY:
                    break
        _connected = status == ROBOTCOM_READY
        if not _connected:
            log('机器人连接未就绪：' + str(msg))
            return False
        RDK.setRunMode(RUNMODE_RUN_ROBOT)
        return True
    except Exception as exc:
        _connected = False
        log('连接失败：' + str(exc))
        return False


# ============================================================
# 解析坐标
# ============================================================
def parse_points():
    if not text_points:
        return []
    raw = text_points.get("1.0", tk.END)
    points = []
    for line in raw.strip().split(NL):
        line = line.strip()
        if not line or line.startswith("#"):
            continue
        try:
            vals = [float(v.strip()) for v in line.split(",")]
            if len(vals) >= 6:
                points.append(vals[:6])
        except ValueError:
            pass
    return points

# ============================================================
# 读取当前位置
# ============================================================
def read_current(entries=None):
    try:
        pose = robot.Pose()
        v = pose_to_fanuc(pose)
        log("")
        log("当前 TCP：X=%.3f Y=%.3f Z=%.3f Rx=%.3f Ry=%.3f Rz=%.3f" % tuple(v[:6]))
    except Exception as e:
        log("读取失败：%s" % e)

def fill_current(entries=None):
    try:
        pose = robot.Pose()
        v = pose_to_fanuc(pose)
        if entries:
            for e, val in zip(entries, v):
                e.delete(0, tk.END)
                e.insert(0, "%.3f" % val)
        log("当前 TCP 已填入")
    except Exception as e:
        log("读取失败：%s" % e)

# ============================================================
# IK 检测
# 注意：SolveIK 显式使用当前 Tool + Reference，和 MoveL/MoveJ 保持一致。
# ============================================================
def check_ik_single(entries=None):
    if not entries:
        return
    try:
        values = [float(e.get()) for e in entries]
    except ValueError:
        log("输入无效")
        return

    x, y, z, rx, ry, rz = values
    target = fanuc_to_pose(x, y, z, rx, ry, rz)
    log("")
    log("目标：X=%.3f Y=%.3f Z=%.3f Rx=%.3f Ry=%.3f Rz=%.3f" % (x, y, z, rx, ry, rz))

    try:
        tool_pose = robot.PoseTool()
        frame_pose = robot.PoseFrame()
        joints = robot.SolveIK(target, tool=tool_pose, reference=frame_pose)
        if joints is None:
            log("IK 不可达")
        else:
            q = joints.list()
            if len(q) < 6:
                log("IK 返回关节数量异常：%d，原始数据=%r" % (len(q), q))
                return
            log("IK 可达")
            log("  关节：J1=%.2f J2=%.2f J3=%.2f J4=%.2f J5=%.2f J6=%.2f" % tuple(q[:6]))
    except Exception as e:
        log("检测失败：%s" % e)

def check_all_ik():
    points = parse_points()
    if not points:
        log("没有有效点")
        return

    log("")
    log("========== 检测全部 %d 个点 ==========" % len(points))
    all_ok = True
    for i, p in enumerate(points):
        try:
            target = fanuc_to_pose(*p)
            joints = robot.SolveIK(target, tool=robot.PoseTool(), reference=robot.PoseFrame())
            if joints is None:
                log("  P%d: 不可达" % (i+1))
                all_ok = False
            else:
                q = joints.list()
                if len(q) < 6:
                    raise ValueError("IK 返回关节数量异常: %d, raw=%r" % (len(q), q))
                log("  P%d: 可达  J1=%.1f J2=%.1f J3=%.1f J4=%.1f J5=%.1f J6=%.1f" % (i+1, *q[:6]))
        except Exception as e:
            log("  P%d: 检测失败 %s" % (i+1, e))
            all_ok = False
    if all_ok:
        log("全部 %d 个点可达" % len(points))
    else:
        log("存在不可达点，执行前整段预检将拒绝不通过的方案")

# ============================================================
# 执行单点
# ============================================================
def execute_single(entries=None, mtype="MoveL"):
    try:
        if not entries:
            return
        values = [float(e.get()) for e in entries]
        _execute_checked_real([dict(type='TCP', values=values)], single_method=mtype)
    except (ValueError, TypeError) as exc:
        log('单点输入无效：' + str(exc))


# ============================================================
# 连续运动：选项卡3直接输入 TCP / 关节点，逐点检查后加入轨迹
# ============================================================
trajectory_records = []
record_text = None
traj_entries = None
traj_type = None
singular_var = None
j6_direction_var = None
spin_var = None


def _parse_six_from_entries(entries, label):
    if not entries or len(entries) != 6:
        log("%s输入框异常：需要 6 个值" % label)
        return None
    try:
        vals = [float(e.get().strip()) for e in entries]
    except (ValueError, AttributeError):
        log("%s输入无效：6 个值必须全部为数字" % label)
        return None
    if not all(math.isfinite(v) for v in vals):
        log("%s输入无效：不能包含 NaN 或无穷值" % label)
        return None
    return vals


def _check_tcp_reachable(vals):
    """检查单个 TCP 点 IK 是否可达，返回 (True, target, joints)。"""
    try:
        target = fanuc_to_pose(*vals)
        tool_pose = robot.PoseTool()
        frame_pose = robot.PoseFrame()
        joints = robot.SolveIK(target, tool=tool_pose, reference=frame_pose)

        if joints is None:
            log("TCP IK：不可达")
            return False, None, None

        q = joints.list()
        if len(q) < 6:
            log("TCP IK：返回关节数量异常：%r" % q)
            return False, None, None

        log("TCP IK：可达")
        log("  IK关节：J1=%.2f J2=%.2f J3=%.2f J4=%.2f J5=%.2f J6=%.2f" % tuple(q[:6]))
        return True, target, q[:6]
    except Exception as e:
        log("TCP IK 检查失败：%s: %s" % (type(e).__name__, e))
        return False, None, None


def _check_tcp_segment_continuous(prev_vals, curr_vals, segment_index, samples=20):
    """检查前一个 TCP 点到当前 TCP 点之间的整段插补路径 IK 连续可达性。

    暂不考虑障碍物，只对 TCP 位姿做线性插值，并对每个采样位姿执行 SolveIK。
    起点和终点也包含在采样检查中。
    """
    if prev_vals is None:
        return True

    log("开始检查 P%d -> P%d 的 TCP 连续 IK（%d 个采样点）" %
        (segment_index - 1, segment_index, samples + 1))

    tool_pose = robot.PoseTool()
    frame_pose = robot.PoseFrame()

    for k in range(samples + 1):
        t = float(k) / float(samples)
        vals = [prev_vals[i] + (curr_vals[i] - prev_vals[i]) * t for i in range(6)]
        try:
            pose = fanuc_to_pose(*vals)
            joints = robot.SolveIK(pose, tool=tool_pose, reference=frame_pose)
            if joints is None:
                log("  P%d -> P%d：第 %d/%d 个采样点 IK 不可达，t=%.3f" %
                    (segment_index - 1, segment_index, k + 1, samples + 1, t))
                log("  TCP：X=%.3f Y=%.3f Z=%.3f Rx=%.3f Ry=%.3f Rz=%.3f" % tuple(vals))
                return False
            q = joints.list()
            if len(q) < 6:
                log("  P%d -> P%d：第 %d 个采样点 IK 返回异常：%r" %
                    (segment_index - 1, segment_index, k + 1, q))
                return False
        except Exception as e:
            log("  P%d -> P%d：第 %d 个采样点 IK 检查失败：%s: %s" %
                (segment_index - 1, segment_index, k + 1, type(e).__name__, e))
            return False

    log("P%d -> P%d：连续 IK 检查通过" % (segment_index - 1, segment_index))
    return True


def _check_joint_reachable(q):
    """兼容旧代码：关节点不做可达性/限位检查，输入合法即可加入。"""
    return True


def refresh_record_list():
    if record_text is None:
        return

    record_text.delete("1.0", tk.END)

    for i, rec in enumerate(trajectory_records, 1):
        kind = rec["type"]
        vals = rec["values"]

        if kind == "TCP":
            if rec.get("spin360", False):
                mark = " [J6自转360° %s]" % ("+" if rec.get("j6_delta", 360) >= 0 else "-")
            elif rec.get("singular", False):
                mark = " [J6特异点 %s180°]" % ("+" if rec.get("j6_delta", 180) >= 0 else "-")
            else:
                mark = ""
            record_text.insert(
                tk.END,
                "P%-3d [TCP]%s   X=%9.3f Y=%9.3f Z=%9.3f Rx=%8.3f Ry=%8.3f Rz=%8.3f%s" %
                (i, mark, *vals, NL)
            )
        else:
            record_text.insert(
                tk.END,
                "P%-3d [JNT]   J1=%8.3f J2=%8.3f J3=%8.3f J4=%8.3f J5=%8.3f J6=%8.3f%s" %
                (i, *vals, NL)
            )


def add_and_check_trajectory_point():
    values = _parse_six_from_entries(traj_entries, traj_type.get())
    if values is None:
        return
    kind = traj_type.get()
    is_singular = kind == 'TCP' and bool(singular_var.get())
    spin = is_singular and bool(spin_var.get())
    sign = 1 if int(j6_direction_var.get()) >= 0 else -1
    rec = dict(type=kind, values=values, singular=is_singular, spin360=spin,
               j6_delta=sign * (360 if spin else 180))
    try:
        records = _validated_records(trajectory_records + [rec])
    except ValueError as exc:
        log('点未加入：' + str(exc))
        return
    trajectory_records[:] = records
    refresh_record_list()
    if spin:
        log('P%d [TCP-J6自转360°]：已加入；执行时 J1~J5 不变，J6 %+d°。' % (len(records), sign * 360))
    else:
        log('点已加入；完整避障预检将在执行前进行。关节圈数按输入保留。')



def _write_values_to_traj_entries(values, label):
    if not traj_entries or len(traj_entries) != 6:
        log("连续运动输入框异常：无法写入当前%s" % label)
        return False
    for e, val in zip(traj_entries, values[:6]):
        e.delete(0, tk.END)
        e.insert(0, "%.3f" % float(val))
    log("当前%s已写入选项卡3输入框" % label)
    return True


def read_current_tcp_to_traj():
    """读取当前 RoboDK TCP，并写入选项卡3的 TCP 输入框。"""
    try:
        pose = robot.Pose()
        vals = pose_to_fanuc(pose)
        log("========== 读取当前 TCP -> 选项卡3 ==========")
        log("X=%+.3f Y=%+.3f Z=%+.3f Rx=%+.3f Ry=%+.3f Rz=%+.3f" % tuple(vals))
        if traj_type.get() != "TCP":
            traj_type.set("TCP")
            _update_traj_labels_and_defaults()
        return _write_values_to_traj_entries(vals, "TCP")
    except Exception as e:
        log("读取当前 TCP 失败：%s: %s" % (type(e).__name__, e))
        return False


def read_current_joints_to_traj():
    """读取 RoboDK Robot Item 当前关节，并写入选项卡3的关节输入框。"""
    q = read_current_joints(None)
    if q is None or len(q) < 6:
        return False
    log("========== 读取当前关节 -> 选项卡3 ==========")
    if traj_type.get() != "JOINT":
        traj_type.set("JOINT")
        _update_traj_labels_and_defaults()
    return _write_values_to_traj_entries(q, "关节")


def clear_trajectory_input():
    if not traj_entries:
        return

    for e in traj_entries:
        e.delete(0, tk.END)

    if traj_type.get() == "TCP":
        defaults = ["0.000", "-241.500", "1047.000", "-90.000", "0.000", "180.000"]
    else:
        defaults = ["0.000"] * 6

    for e, val in zip(traj_entries, defaults):
        e.insert(0, val)




def import_trajectory():
    filepath = filedialog.askopenfilename(title='导入轨迹', defaultextension='.json', filetypes=[('JSON轨迹','*.json'),('所有文件','*.*')])
    if not filepath:
        return
    try:
        with open(filepath, encoding='utf-8') as f:
            records = _validated_records(json.load(f))
        trajectory_records[:] = records
        refresh_record_list()
        log(f'已导入{len(records)}点：{filepath}。执行前将从实机当前关节重新预检。')
    except Exception as exc:
        log('轨迹导入失败：' + str(exc))


def delete_last_record():
    if trajectory_records:
        rec = trajectory_records.pop()
        refresh_record_list()
        log("已删除最后一点：P%d [%s]" %
            (len(trajectory_records) + 1, rec["type"]))
    else:
        log("当前没有可删除的连续运动点")


def clear_records():
    trajectory_records.clear()
    refresh_record_list()
    log("连续运动点列表已清空")


def execute_recorded_trajectory():
    log('【点击】执行整段连续运动：当前列表 %d 点（转后台线程执行，窗口保持响应）' % len(trajectory_records))
    import threading
    def _worker():
        try:
            _execute_checked_real(list(trajectory_records))
        except Exception as exc:
            log('【线程异常】%s: %s' % (type(exc).__name__, exc))
    threading.Thread(target=_worker, daemon=True, name='real_exec').start()



# 保留旧函数名，避免其他代码调用失效。
def execute_trajectory():
    execute_recorded_trajectory()


# ============================================================
# 实机关节运动
# ============================================================
def _joint_values_from_entries(entries):
    """从 GUI 读取 J1~J6 目标角度。单位：deg。"""
    if not entries or len(entries) != 6:
        log("目标关节输入框异常：需要 J1~J6 共 6 个")
        return None
    try:
        q = [float(e.get().strip()) for e in entries]
    except (ValueError, AttributeError):
        log("目标关节输入无效：J1~J6 必须全部填写数字")
        return None
    if not all(math.isfinite(v) for v in q):
        log("目标关节输入无效：不能包含 NaN 或无穷值")
        return None
    return q


def read_current_joints(entries=None):
    """读取 RoboDK Robot Item 当前关节值，并可直接填入 J1~J6 输入框。
    注意：这里读取的是 RoboDK 当前 Robot Item 的关节状态，不调用 CR5 控制器 GetAngle。
    """
    try:
        joints = robot.SimulatorJoints()
        q = list(joints) if hasattr(joints, "__iter__") else [joints]
        if len(q) < 6:
            log("读取当前关节失败：SimulatorJoints 返回 %r" % (q,))
            log("请确认 RoboDK 窗口中的机器人已经连接并显示实时关节角度。")
            return None

        q = q[:6]
        log("")
        log("========== RoboDK 当前关节 ==========")
        log("J1=%+.3f°  J2=%+.3f°  J3=%+.3f°" % tuple(q[:3]))
        log("J4=%+.3f°  J5=%+.3f°  J6=%+.3f°" % tuple(q[3:]))

        if entries and len(entries) == 6:
            for e, val in zip(entries, q):
                e.delete(0, tk.END)
                e.insert(0, "%.3f" % val)
            log("当前关节已填入 J1~J6 输入框")

        return q
    except Exception as e:
        log("读取 RoboDK 当前关节失败：%s: %s" % (type(e).__name__, e))
        return None


def fill_current_joints(entries=None):
    """当前 RoboDK 关节 -> 目标关节输入框。"""
    return read_current_joints(entries)


def execute_joint_target(entries=None):
    q = _joint_values_from_entries(entries)
    if q is not None:
        _execute_checked_real([dict(type='JOINT', values=q)])



def clear_joint_target(entries=None):
    if not entries:
        return
    for e in entries:
        e.delete(0, tk.END)
        e.insert(0, "0.000")
    log("目标关节输入已清零")

# ============================================================
# GUI
# ============================================================

# 与TCP仿真一致的预检核心；仅在仿真模式调用。
fanuc_values_to_pose = fanuc_to_pose
pose_to_fanuc_values = pose_to_fanuc
MOVEJ_FALLBACK_MAX_DEVIATION_MM = 50.0
# 预检缓存（与TCP仿真副本同款）：生命周期=单次预检规划，_enable_obstacle_checks 每次进入预检时清空。

_plan_cache = {}
_preferred_seed = None  # Ordering hint only; never reuse a collision certificate.


def _lazy_valid_seeds(seeds, start):
    """Keep the existing valid-seed order, testing only seeds actually needed.

    If none is reachable, preserve the old fallback to the unfiltered list.
    """
    found = False
    for seed in seeds:
        if seed is None or _movej_test_cached(start, seed, 1) == 0:
            found = True
            yield seed
    if not found:
        yield from seeds

def _cache_key_joints(q):
    return tuple(round(float(v), 3) for v in q[:6])

def _cache_key_pose(pose):
    return tuple(tuple(round(float(v), 6) for v in row) for row in pose.rows)

def _movej_test_cached(start, end, minstep_deg):
    """robot.MoveJ_Test 的缓存包装，返回值与直接调用完全一致。
    成功时与原调用一样把仿真关节停在终点；失败路径的规划器只依赖局部
    关节变量（不读取此时的模型关节状态），无需复现失败的副作用。"""
    key = ('movej_test', _cache_key_joints(start), _cache_key_joints(end),
           round(float(minstep_deg), 6))
    if key not in _plan_cache:
        _plan_cache[key] = robot.MoveJ_Test(start, end, minstep_deg=minstep_deg)
    elif _plan_cache[key] == 0:
        robot.setJoints(list(end[:6]))
    return _plan_cache[key]

def _tcp_target_to_flange(target):
    """输入是参考系中的TCP；IK需要机器人基座系中的法兰位姿。"""
    return robot.PoseFrame() * target * invH(robot.PoseTool())

def _flange_target_description(target):
    flange = _tcp_target_to_flange(target)
    return ('换算后的法兰中心（基座系）XYZ=' +
            str(tuple(round(v, 3) for v in flange.Pos())) +
            ' mm，法兰Z轴方向=' + str(tuple(round(v, 6) for v in flange.VZ())))


def _validated_records(data):
    if not isinstance(data, list) or not data:
        raise ValueError('轨迹必须是非空点列表。')
    result = []
    for i, rec in enumerate(data, 1):
        kind = str(rec.get('type', '')).upper()
        if kind == 'JNT':
            kind = 'JOINT'
        values = [float(v) for v in rec.get('values', [])]
        if kind not in ('TCP', 'JOINT') or len(values) != 6 or not all(math.isfinite(v) for v in values):
            raise ValueError(f'P{i}：类型或六维数值无效。')
        special = bool(rec.get('singular', False)) and kind == 'TCP'
        spin = special and bool(rec.get('spin360', False))
        raw_delta = int(rec.get('j6_delta', 360 if spin else 180)) if special else 0
        if special and (not result or result[-1]['type'] != 'TCP' or result[-1]['singular']):
            raise ValueError(f'P{i}：特异点前序或转向无效。')
        if special:
            if spin:
                if raw_delta not in (-360, 360):
                    raise ValueError(f'P{i}：J6自转方向必须为+360或-360。')
                if max(abs(a - b) for a, b in zip(values, result[-1]['values'])) > 1e-3:
                    raise ValueError(f'P{i}：J6自转360°特异点的六维数值必须与前一个TCP点完全相同。')
            elif raw_delta not in (-180, 180):
                raise ValueError(f'P{i}：J6方向必须为+180或-180。')
        delta = (360 if spin else 180) * (1 if raw_delta >= 0 else -1) if special else 0
        result.append(dict(type=kind, values=values, singular=special, spin360=spin, j6_delta=delta))
    return result


def _controller_feedback():
    # Dobot CR V3: 1440-byte real-time feedback; no command is sent on this socket.
    import socket
    import struct
    host, port, *_ = robot.ConnectionParams()
    if int(port) != 29999:
        raise RuntimeError('当前连接不是已验证的Dobot CR反馈协议。')
    previous = None
    with socket.create_connection((host, 30004), timeout=3.0) as connection:
        deadline = time.monotonic() + 3.0
        for _ in range(2):
            packet = bytearray()
            while len(packet) < 1440:
                remaining = deadline - time.monotonic()
                if remaining <= 0:
                    raise RuntimeError('实机反馈读取超时。')
                connection.settimeout(remaining)
                part = connection.recv(1440 - len(packet))
                if not part:
                    raise RuntimeError('实机反馈连接已关闭。')
                packet.extend(part)
            length = struct.unpack_from('<Q', packet, 0)[0]
            marker = struct.unpack_from('<Q', packet, 48)[0]
            stamp = struct.unpack_from('<Q', packet, 32)[0]
            if length != 1440 or marker != 0x123456789ABCDEF:
                raise RuntimeError('实机反馈帧格式不匹配。')
            if previous is not None and stamp <= previous:
                raise RuntimeError('实机反馈时间戳未更新。')
            previous = stamp
        q = list(struct.unpack_from('<6d', packet, 192))   # ★真实关节角（v10定位，示教器交叉证实）；旧版误读432="连接基准+指令累加"的假值
        velocity = list(struct.unpack_from('<6d', packet, 480))
        mode = struct.unpack_from('<Q', packet, 24)[0]
        if not all(math.isfinite(v) for v in q + velocity):
            raise RuntimeError('实机反馈包含无效关节数值。')
        return q, velocity, mode


def _live_joints():
    if RDK.RunMode() != RUNMODE_RUN_ROBOT:
        raise RuntimeError('当前不是实机执行模式。')
    status, msg = robot.ConnectedState()
    if status != ROBOTCOM_READY:
        raise RuntimeError('机器人未就绪或已断连：' + str(msg))
    q, velocity, mode = _controller_feedback()
    # 阈值由 0.1 放宽到 1.0：实测静止时 J4/J3 的速度估计噪声可达 0.31°/s
    # （六轴角度 8 次采样完全相同），0.1 会把"其实已静止"误判为运动中而中止任务。
    if mode != 5 or max(abs(v) for v in velocity) > 1.0:
        raise RuntimeError('实机未处于使能静止状态，模式=%s。' % mode)
    return q


def _require_joints(expected, _tries=3, _allow_fix=False):
    """校验关节与预检一致（容差 0.5°）；失败时【主动发一条 MoveJ 校正】，仍不行才抛错。

    ★★★ v15.10（2026-11-03）：根治"走到 P8 后不动"。
    根因（读码确认）：`_settle_core` 的断连分支写的是
        `_wait_arrival_then_static(expect_target)`
      · 直发段传了 expect_target ⇒ 会等到目标 ✓
      · **MoveJ 段传的是 None** ⇒ 退化为「只等静止」✗
      ⇒ 指令被断连打断、手臂停在中途 ⇒ 只要「静止」就算完成 ✗
      ⇒ 下一段开头的 _require_joints 发现差 9.77° ⇒ 抛错 ⇒ 停 ✗
    （历史证据：10-13 12:12 / 15:49 / 15:55 三次同样失败，当时 P8 走的是纯 MoveJ，与直发无关 ✗）

    修法：不再是"发现不一致就停"，而是【发一条 MoveJ 到认证关节】把手臂拉回去，再校验。
      · 目标就是预检认证过的关节构型 ⇒ 确定可达 ⇒ 重发安全 ✓
      · 只补一次（_allow_fix=False 时不再递归）⇒ 不会无限循环 ✓
      · 拉回后仍不一致 ⇒ 才抛错 ✓（护栏不放松）
    """
    last = None
    actual = None
    for k in range(_tries):
        actual = _live_joints()
        last = max(abs(a - b) for a, b in zip(actual, expected))
        if last <= 0.5:
            return
        if k < _tries - 1:
            log('关节偏差 %.2f° > 0.5°（第 %d/%d 次）⇒ 等 0.5s 重读（可能仍在微动）'
                % (last, k + 1, _tries))
            time.sleep(0.5)
    if _allow_fix:
        log('关节偏差 %.2f°（目标%s，实测%s）⇒ 主动发 MoveJ 校正到认证关节（v15.10）'
            % (last, ['%.2f' % v for v in expected], ['%.2f' % v for v in (actual or [])]))
        try:
            robot.MoveJ(list(expected))
            time.sleep(1.0)
            _require_joints(expected, _tries=3, _allow_fix=False)
            log('✓ 校正 MoveJ 生效：关节已回到认证构型')
            return
        except Exception as _fix_exc:  # noqa: BLE001
            log('⚠️ 校正 MoveJ 未生效：%s: %s' % (type(_fix_exc).__name__, _fix_exc))
    raise RuntimeError('关节反馈与预检状态不一致（偏差 %.2f°，目标%s，实测%s），停止后续命令。'
                       % (last, ['%.2f' % v for v in expected], ['%.2f' % v for v in (actual or [])]))


def _retreat_orientation_records(records):
    """加工点变姿态前退到 y=-750，变姿态后返回 y=-775。"""
    result = []
    previous = None
    for index, record in enumerate(records, 1):
        current = dict(record, values=record['values'][:])
        current['label'] = f'P{index}'
        if previous and previous['type'] == current['type'] == 'TCP':
            old, new = previous['values'], current['values']
            changed = pose_angle(invH(fanuc_values_to_pose(*old)) * fanuc_values_to_pose(*new)) > math.radians(.01)
            old_work, new_work = abs(old[1] + 775) < .001, abs(new[1] + 775) < .001
            if changed and (old_work or new_work):
                anchor = old if old_work else new
                retreat = dict(type='TCP', values=[anchor[0], -750., anchor[2]] + old[3:], singular=False,
                               label=f'P{index}前退让', require_linear=old_work)
                result.append(retreat)
                turn = dict(current, values=retreat['values'][:3] + new[3:], label=f'P{index}退让位换向')
                result.append(turn)
                current['singular'] = False
                current['require_linear'] = new_work
        result.append(current)
        previous = record
    return result


def _prepare_real_plan(records, start, deviation, single_method=None):
    RDK.setRunMode(RUNMODE_SIMULATE)
    try:
        RDK.Command('Trace', 'Off')
        robot.setJoints(start)
        if single_method is None:
            return _plan_continuous_trajectory(records, deviation, log)
        _enable_obstacle_checks()
        if robot.MoveJ_Test(start, start, minstep_deg=1) != 0:
            raise ValueError('起始姿态碰撞：' + _collision_details())
        values = records[0]['values']
        method, fallback = single_method, False
        if method not in ('MoveJ','MoveL'):
            raise ValueError('未知单点运动类型。')
        end = None
        waypoints = []
        if method == 'MoveL':
            end, _ = _linear_path_endpoint(start, fanuc_to_pose(*values))
            if end is not None:
                # v13：单点 MoveL 同样不信任驱动 MOVL（纯J6自转也一样，关节插值=同一路径），
                # 改细分途经点+MoveJ 执行
                waypoints = _linear_waypoints(start, fanuc_to_pose(*values))
                if waypoints:
                    log('单点 MoveL 改细分执行：%d 个途经点（步长≤%.0fmm）。' % (len(waypoints), LINEAR_SUBSTEP_MM))
                    log('单点 MoveL 途经跳（共%d跳）：%s' % (len(waypoints), [[float('%.2f' % v) for v in w] for w in waypoints]))
        if end is None:
            end = _obstacle_joint_target(start, values, deviation if method=='MoveL' else None)
            fallback, method = method=='MoveL', 'MoveJ'
        plan = [dict(method=method,joints=end,special=False,fallback=fallback,rewinds=[],j6_delta=None,waypoints=waypoints)]
        _verify_obstacle_plan(start, plan)
        return plan
    finally:
        robot.setJoints(start)
        RDK.Render(True)
        RDK.setRunMode(RUNMODE_RUN_ROBOT)  # 旧版 L615 有此行：预检后必须切回实机模式，否则 _live_joints 直接拒执行


def _wait_controller_static(max_wait_s=20.0, vel_threshold=0.5, samples=5, interval=0.3):
    """轮询30004反馈直到六轴静止（连续samples次速度<阈值），返回(关节, 是否静止)。

    v14o：断连分支以 samples=3/interval=0.2 调用（短跳≈1s，5×0.3s 静止确认占每跳
    尾部 ~1.5s，是停顿税大头）；默认 5×0.3s 供正常路径；20s 静止上限（真断连护栏）不动。"""
    t0 = time.time()
    quiet = 0
    last = None
    while time.time() - t0 < max_wait_s:
        actual, velocity, _mode = _controller_feedback()
        last = actual
        if max(abs(v) for v in velocity) < vel_threshold:
            quiet += 1
            if quiet >= samples:
                return last, True
        else:
            quiet = 0
        time.sleep(interval)
    return last, False


class ControllerMotionFault(RuntimeError):
    """A controller state that must never trigger a motion resend."""
    pass


def _wait_arrival_then_static(target_joints, max_wait_s=20.0):
    """v14u：目标锚定的到位等待——直发后不再猜「起步了没」，只等「到没到」。

    背景（v14t 10:38 P9 实测）：直发指令起步延迟可 >6s，让位 6s 耗尽判「未执行」
    停止后，指令仍被控制器自行执行到精确目标（善后实测 J2 +10°/J3 +20°，余轴不动，
    宏未重发）——「起点静止」与「完成静止」在反馈上不可区分，位置对目标才是唯一
    可靠锚点（速度判据出局：三场停时 J4 0.06~0.42°/s 均为低于阈值的保持抖动）。
    本函数：距目标关节 ≤MOVL_ARRIVE_TOL_DEG 且速度<0.5°/s → 到位完成（此时已在
    目标，无需再做常规静止确认）；每 5s 一行进度日志（顺带实测真实延迟）；
    上限 MOVL_ARRIVE_WAIT_S 超时报「疑似未执行」停待判读；不重发铁律不变。
    target_joints=None → 退化为 _wait_controller_static()，行为与原先完全一致。"""
    if target_joints is not None:
        t0 = time.time()
        t_note = t0
        while True:
            fb = _controller_feedback()
            if fb[2] not in (5, 7, 8):
                raise ControllerMotionFault(
                    '控制器反馈模式=%s，停止等待且不补发；目标关节=%s，实际关节=%s。请检查示教器报警。'
                    % (fb[2], target_joints, fb[0]))
            err = max(abs(a - b) for a, b in zip(fb[0], target_joints))
            if err <= MOVL_ARRIVE_TOL_DEG and max(abs(v) for v in fb[1]) < 0.5:
                log('MovL 直发到位确认：距目标关节%.2f°（%.1fs），验收继续。'
                    % (err, time.time() - t0))
                return fb[0], True
            if time.time() - t0 >= MOVL_ARRIVE_WAIT_S:
                raise RuntimeError(
                    'MovL 直发%.0fs仍未到位（距目标关节%.2f°），疑似未执行，停止待判读。'
                    % (MOVL_ARRIVE_WAIT_S, err))
            if time.time() - t_note >= 5.0:
                log('MovL 直发等待到位：%.0fs，距目标关节%.2f°，续等（不重发，上限%.0fs）。'
                    % (time.time() - t0, err, MOVL_ARRIVE_WAIT_S))
                t_note = time.time()
            time.sleep(0.5)
    return _wait_controller_static(max_wait_s=max_wait_s)


MOVE_OFFSET_TOL = 0.5   # 闭环补偿后的到位容差（°）


TCP_TOOL_NAME = 'CR5_TCP_130mm'
FLANGE_TOOL_NAME = '_CR5_FLANGE_DIRECT_TEMP'
_tool_window_depth = 0


def _same_tool_pose(a, b):
    return max(abs(a[r, c] - b[r, c]) for r in range(4) for c in range(4)) < 1e-7


def _named_tool(name, pose):
    matches = [it for it in robot.Childs()
               if it.Type() == ITEM_TYPE_TOOL and it.Name() == name]
    if len(matches) > 1:
        raise RuntimeError('重复 TCP 工具条目：' + name)
    if matches:
        tool = matches[0]
        if not _same_tool_pose(tool.PoseTool(), pose):
            raise RuntimeError('TCP 工具定义不符，停止待核对：' + name)
        return tool
    return robot.AddTool(pose, name)


def _restore_tool(pose, linked_tool=None):
    """Restore the original item link when possible, and never swallow failure."""
    for attempt in range(2):
        try:
            robot.setPoseTool(linked_tool if linked_tool is not None and linked_tool.Valid() else pose)
            if not _same_tool_pose(robot.PoseTool(), pose):
                raise RuntimeError('PoseTool 恢复后读回不一致')
            return
        except Exception as exc:
            if attempt == 1:
                raise RuntimeError('工具恢复失败，禁止继续运动：' + str(exc)) from exc


def _single_move_settle(method, target, require_joints=True, expect_target=None, flange_space=False, _retry=0):
    """发指令并确认到位——v14w39 窗口版入口：flange_space 时单位变换+藏把手覆盖
    【整个 settle 生命周期】（发送+断连恢复+到位等待）。旧版只包 RPC 一次调用：假断连
    抛出时窗口即关、把手提前回来，RoboDK 本地退化动画在弧 66% 被碰撞检测掐停→模型冻在
    撞点、红显常驻→收口 MoveJ 被拦死（10-22 四次实录含 v14w38）。"""
    global _tool_window_depth
    if not flange_space or _tool_window_depth:
        # A controlled retry already runs inside the outer tool window.
        # Only the outer owner may restore the original TCP.
        return _settle_core(method, target, require_joints, expect_target, flange_space, _retry)
    _ensure_canonical_tool()
    _win_tp = robot.PoseTool()
    _win_link = robot.getLink(ITEM_TYPE_TOOL)
    _win_handle = RDK.Item('门把手_bs1')
    _win_visible = _win_handle.Visible() if _win_handle.Valid() else None
    _flange_tool = _named_tool(FLANGE_TOOL_NAME, eye(4))
    _tool_window_depth += 1
    try:
        robot.setPoseTool(_flange_tool)
        if not _same_tool_pose(robot.PoseTool(), eye(4)):
            raise RuntimeError('法兰工具切换失败，未发送运动指令')
        if _win_visible is not None:
            _win_handle.setVisible(False)
        result = _settle_core(method, target, require_joints, expect_target, True, _retry)
        # Synchronize measured joints before restoring the tool and visible mesh.
        actual, is_static = _wait_controller_static()
        if not is_static:
            raise RuntimeError('法兰直发后未确认静止，停止后续命令。')
        robot.setJoints(actual)
        return result
    finally:
        try:
            _restore_tool(_win_tp, _win_link)
        finally:
            _tool_window_depth -= 1
            if _win_visible is not None:
                _win_handle.setVisible(_win_visible)


def _settle_core(method, target, require_joints, expect_target, flange_space=False, _retry=0):
    """发一条运动指令并确认到位（v10：反馈字段已校正）。

    v14r：require_joints=False 仅供 MovL 直发调用点使用——断连分支的关节级 0.5°
    校验让位给外层法兰级粗验收（≤8mm/≤1°）+MoveJ 微纠偏收口（v14q 09:57 实机
    教训：MovL 直发必触发假断连，0.95° 固有残差在断连分支内即被拦停，外层验收
    根本没执行到）。其余护栏不变：20s 静止上限、重连失败仍停。

    v14u：断连分支改目标锚定到位等待 _wait_arrival_then_static——上限 60s 每 5s
    进度日志；超时报「疑似未执行」停。不重发铁律不变。

    v14w37：直发=【法兰位姿传递 + flange_space 单位变换窗口】双件套——
    ①传位姿（调用方 invH(PoseFrame)*SolveFK(净化关节) 自算）：MoveL 的动画按位姿空间
    直线走=认证路径，根治旧 MoveL(关节) 的关节弧动画扫进圆柱假碰撞冻死（10-22 两次实录）；
    ②发送 RPC 窗口内 PoseTool 置单位变换：MoveL(位姿) 的可达校验/语义都按 TCP 空间做，
    不切工具则法兰位姿被当 TCP 反推（P8 反推法兰 z=744 爆臂展 ⇒ TargetReachError，
    10-22 11:18 实录）；单位变换下校验空间=法兰空间，数字逐位=金标准（实证 0 偏差）。
    动画窗口内直线途经点 12/12 无碰撞（单位变换工具下实测）。
    v14w38：窗口内追加隐藏把手——驱动断连瞬间 RoboDK 本地退化关节动画（会撞圆柱的
    那条弧）是三次冻结的真凶；藏把手=对假路径的检测放行（实测弧中点/冻结姿态
    显隐 True/False 翻转），真直线 1mm 检查本来就 0 碰撞。

    v14w20：受控补发（一次性）——驱动连接恰死在发送时刻时 SendJointMovJ 会静默
    丢弃不发送（反汇编：CONNECTED=False 直接 return False；2026-10-15 09:51 P25
    实发：断连后臂停在发送前位置、误差127.8°）。补发条件（全部满足才补，且全程
    至多一次）：①失败 ②30004 独立反馈证明【零位移】（仍在发送前关节 ≤0.5°）
    ③ensure_connected() 重连成功。指令已上线/延迟执行/落点异常的场景均不满足
    ②（有位移）不会触发——保留原「不重发」语义。历史上"晚执行"案例（v14t）
    后经控制器日志证实为面板拖动误判，非队列延迟。

    历史结论：驱动一直正确执行绝对关节目标；真实关节角在偏移192。"""
    try:
        _start_q = None
        try:
            _start_q = _controller_feedback()[0]
        except Exception:
            _start_q = None
        getattr(robot, method)(target)   # v14w39：flange 窗口已上移至 _single_move_settle 包装层
    except StoppedError as exc:
        if str(exc).strip() != 'Robot not connected':
            raise
        # v14o 静默重连：假断连是本环境常态（每条 MoveJ 指令结束后都可能误报）；30004
        # 反馈通道独立于驱动连接，静止确认与重连并行进行，压缩跳间停顿税。
        # 护栏不变：未自然收尾（20s 上限）仍停、落点仍 0.5° 校验、重连失败仍停。
        log('驱动报断连——等待收尾与后台重连并行进行…')
        import threading as _st
        reconnected = []
        def _bg_reconnect():
            for _r in range(3):
                if ensure_connected():
                    reconnected.append(True)
                    return
                time.sleep(1.0)
        _rt = _st.Thread(target=_bg_reconnect, daemon=True, name='silent_reconnect')
        _rt.start()
        # v14u：到位等待下沉在断连分支（MovL 直发永远走本分支——v14s 教训）——
        # 目标锚定：距目标≤2°且静止=完成，不猜起步。非 MovL 直发退化为常规静止确认。
        try:
            actual, is_static = _wait_arrival_then_static(expect_target)
        except RuntimeError as _arr_exc:
            if isinstance(_arr_exc, ControllerMotionFault):
                raise
            # v14w20：直发「疑似未执行」——零位移+重连成功 ⇒ 补发一次（指令未上线实证）
            if (_retry < 1 and _start_q is not None
                    and max(abs(a - b) for a, b in zip(_controller_feedback()[0], _start_q)) <= MOVE_OFFSET_TOL
                    and ensure_connected()):
                log('直发疑似未执行且零位移（仍在起点）——判定指令未上线，补发一次（v14w20）。')
                return _single_move_settle(method, target, require_joints, expect_target,
                                           flange_space, _retry=_retry + 1)
            raise
        if not is_static:
            raise RuntimeError('驱动报断连后等待%.0fs仍未静止，停止。' % 20.0) from exc
        if require_joints:
            err = max(abs(a - b) for a, b in zip(actual, target))
            if err > MOVE_OFFSET_TOL:
                # v14w20：MoveJ 类「断连收尾后未到位」——零位移+重连成功 ⇒ 补发一次
                if (_retry < 1 and _start_q is not None
                        and max(abs(a - b) for a, b in zip(actual, _start_q)) <= MOVE_OFFSET_TOL
                        and ensure_connected()):
                    log('断连后零位移（仍在起点）——判定指令未上线，补发一次（v14w20）。')
                    return _single_move_settle(method, target, require_joints, expect_target,
                                               flange_space, _retry=_retry + 1)
                raise RuntimeError('断连收尾后未到位：目标%s，实测%s（误差%.2f°），停止待判读。'
                                   % (['%.2f' % v for v in target], ['%.2f' % v for v in actual], err)) from exc
        _rt.join(timeout=4.0)
        if not reconnected:
            raise RuntimeError('已到位但驱动重连失败，停止后续指令。') from exc
        log('驱动断连但运动已自然完成到位；已重连驱动，继续。')
        return
    actual, is_static = _wait_controller_static()
    if not is_static:
        raise RuntimeError('指令返回后等待静止超时（20s），停止。')
    if require_joints:
        err = max(abs(a - b) for a, b in zip(actual, target))
        if err > MOVE_OFFSET_TOL:
            raise RuntimeError('落点偏差%.2f°：目标%s，实测%s，停止待判读。'
                               % (err, ['%.2f' % v for v in target], ['%.2f' % v for v in actual]))
    return


MOVE_OFFSET_TOL = 0.5   # 到位容差（°）：反馈字段校正后，超过即停止待判读


# v13（方案B）：驱动 MOVL 执行层已判死（3 次实机断连指纹 + .pyc 反汇编直连无收尾），
# 所有 MoveL 执行全部替换为「细分途经点 + MoveJ」。作业面短段（≤ TRANSIT_DIRECT_MAX_MM）
# 用 MoveL 指令的 1mm 逆解采样出 ≤ LINEAR_SUBSTEP_MM 的途经关节序列，MoveJ 逐跳执行；
# 过渡段长段优先 MoveJ 直达（须过 TCP 偏离≤max_deviation 且整弧 MoveJ_Test 碰撞检查），
# 不满足才退回细分。预检层 MoveL_Test@1mm 保留：仍是「这一段能不能走直线」的权威筛选器。
TRANSIT_DIRECT_MAX_MM = 300.0   # 超过此段长的 TCP 段视为自由空间过渡段，尝试 MoveJ 直达
LINEAR_SUBSTEP_MM = 20.0        # 作业面细分步长：v14m(40mm) 实机碰撞实证弦误差可吃掉真裕度（轴线距199.9-半径180≈19.9mm），回 20mm 安全基准（v14k 两度全通过）；途经点弦误差 <0.5mm

MOVL_DIRECT_MAX_MM = 250.0   # v14w35（10-22）：150→210——150 是 v14p 照当时谱系（最长≈120mm）取的设计余量，非事故判死值；210 覆盖 200mm 工艺段一指令（y=-719 线翻转点→x=-100），留 FP 边界余量。路径背书不变（认证直线+整段复核）；更长直线段仍走细分
# ★★★ v14w（2026-10-13 16:08）：【禁直发名单清空 = 恢复 P9 直发】+ 发送位姿数字净化。
#   v14v4 按点号拦 P9 是在 -30001 真凶查明前的临时措施（且拦下分支会落空——随名单清空，
#   该落空分支变为不可达死码，留档不删）。真凶 = 控制器 MovL 参数校验拒收【参数形态】
#   （-0.000000 / +90.000000 / -0.000000，见 LOG_VERSION 处实录），不是几何、不是段长：
#   同目标 15:55:51 单步直发实证 return 0、1.1s 到位。净化失败 ⇒ 本段自动改走细分（安全回落）。
# 想再拦某点：改回 (9,) 即可（注意拦下分支的落空缺陷仍在，见 P2P_LESSONS.md）。
# ★★★ 2026-11-03：改回 (9,) —— 针对【新根因】"movL not set tool or user"（不是 -30001）
#   实录（控制器日志 11-03 10:33:24 / 10:33:30）：
#     [MovL#859] Motion args is legal!            ← 参数合法（所以不是 -30001）
#     [MovL#878] movL not set tool or user!!!     ← ★ 工具/用户坐标系没设置
#     [CallProcess#275] ret = 73/76 ... return = 0,{}  ← 被接受，但按【默认 tool/user】执行
#   ⇒ RoboDK 的 DobotCR 驱动下发 MovL(x,y,z,rx,ry,rz) 时【不带 tool/user】✗
#     ⇒ 控制器用开机默认值 ⇒ 与脚本"法兰补偿（PoseTool=eye）"的语义不一致 ⇒ 落点偏离（P9 差 11.80°）✗
#   ⇒ 保底：P9 不做直发，直接走【细分途经点路径】（今天 P5 就是这样走完的：13 途经点 ✓）
#   ⇒ 根治手段见下方 MOVL_SEND_TOOL_USER（实验性，默认关）
# ★★★ v15.9（2026-11-03）：P8 也加入禁直发 —— 直发的"选解自由"问题对 P8 同样致命。
#   实录（v15.8, 11:56:09~14）：
#     P8 直发 → 等静止 ✓ → 法兰验收通过（5.71mm/0.32° ✓）→ 收口 MoveJ
#     ⇒ 控制器最后停在【另一组 IK 解】：
#        目标 [68.33, 41.30, 10.92, 37.78, -90, 158.33]
#        实测 [78.10, 36.86, 19.48, 33.66, -90, 168.10]
#        差   +9.77, -4.44, +8.56, -4.12,  0,  +9.77
#     ⇒ J1 与 J6 同步 +9.77° ⇒ 【基座-腕部互相补偿】的同一法兰位姿、另一组解 ✗
#   ⇒ 根因：MovL 只给位姿 ⇒ 控制器自行选 IK 分支 ⇒ 关节构型不可控 ✗
#     （v15.5~v15.8 的等待/重试/安全网都改变不了这一点 ✗）
#   ⇒ 细分路径是【逐关节】走的 ⇒ 不存在选解问题 ⇒ 关节精确 ✓（代价：8 跳 ≈24 秒）
MOVL_DIRECT_BLOCK_POINTS = (9, 11)

# ★ 实验性开关（v15.3 已打开做验证）：直发前先给【控制器】发 Tool(0)/User(0)，
#   让 MovL 明确用 基座系+零工具(法兰)。背景：[MovL#878] movL not set tool or user!!!
#   ⇒ 控制器没收到 tool/user 就按默认执行 ⇒ 与"法兰补偿（PoseTool=eye）"语义不一致 ⇒ P9 落点偏 11.80°
#   验证目标：打开后控制器日志里 `movL not set tool or user` 是否消失。
#     消失 ⇒ 直发侧真能用 ⇒ "断断续续"（13 跳 × 3 秒）可根治 ✓
#     仍出现 ⇒ RoboDK DobotCR 驱动不透传 Tool()/User() ⇒ 此路不通，只能接受 3 秒/跳 ✗
#   安全性：发送失败只记日志、不阻断主流程；直发落点仍受法兰级粗验收（≤8mm/≤1°）护栏 ✓
MOVL_SEND_TOOL_USER = False  # RunCodeCustom is a project call, not raw dashboard transmission.
MOVL_FLANGE_TOL_MM = 8.0     # v14q 直发 MovL 法兰位置粗验收容差：控制器 MovL 固有落点残差实测 4.61mm（v14p 首航）/5.5mm（v14l）双样本，取实测+裕量；超此值=落点异常真停
MOVL_FLANGE_TOL_DEG = 1.0    # v14q 直发 MovL 法兰姿态粗验收容差（实测 0.616°+裕量）；通过后 MoveJ 微纠偏收口到关节级 0.5° 内
MOVL_ARRIVE_WAIT_S = 60.0    # v14u MovL 直发到位等待上限：目标锚定（距目标≤2°且静止即完成），不猜起步——v14t 10:38 实测 P9 起步延迟>6s、指令事后自行执行完；60s 为 10 倍裕量，每5s进度日志实测真实延迟，超时按未执行停待判读
MOVL_ARRIVE_TOL_DEG = 5.0    # v14u 到位判定关节距离阈（°）；v14w30 2→5：tool=182 构型下 ~5mm 固有误差映射关节达 2.58°（10-21 P8 实证），阈外即误判未执行——粗验收前哨放宽，法兰级粗验收(≤8mm/≤1°)+MoveJ收口紧随其后罩终点；此处不走 MOVE_OFFSET_TOL=0.5°（require_joints=False 路径，护栏语义不降级）

# v14w22：实机关节限位（与 RoboDK 模型 ±360 取交集）。依据：J1=193.59 两次被控制器
# -40001 拒收（10-15 P25）；J6=190.84 return 0 ✓；J5=177.6 实机走成 ✓（故 J5=180 非
# 某些资料的 ±120）；J3 取模型更紧的 ±160。规划期过滤，保证预检路径=实发路径。
# v14w23：J4 190→150——J4=-189.70 被控制器 -40004（自干涉 PoseSelfInterference）拒收；
# -168 族中途自干涉保护停机；实证安全族 |J4|≤95，150 留 55° 余量。
# ★★★ 2026-11-03：J4 150→178（用户要求）★★★
#   原因：150 太紧 ⇒ 某些点的【全部 IK 解都被过滤】⇒ 报 "ValueError: 没有限位内的逆解"
#         （11-03 10:29:35 实测：已完成 0 点即停）。要让那些点出解，J4 必须 ≥165。
#   代价：(150,178] 区间【重新暴露 -40004 自干涉拒收】风险 ✗
#         ⇒ 依靠 REAL_INTERFERE_J4_MAX / REAL_INTERFERE_J5_MIN（J4×J5 组合区禁选）
#           + 规划期预检（MoveJ_Test / MoveL_Test）兜底；
#         ⇒ 若再现 -40004，把本值在 165~178 之间微调（165 = "能出解 + 少踩禁区"的折中）。
#   历史：190 ✗(-40004) → 150 ✓（安全但出解困难）→ 178（本次，兼顾出解）
REAL_JOINT_LIMITS = (180.0, 180.0, 160.0, 178.0, 180.0, 360.0)

# v14w26：实机自干涉组合区（控制器 PoseSelfInterference 的 J4×J5 耦合，-40006）。
# 实录：|J4|=115.5×|J5|=173.1 与 |J4|=109.4×|J5|=171.5 均拒；|J4|=83.2×|J5|=177.6 通过。
# 阈值取中：|J4|>100 且 |J5|>165 视为禁区（两端各留 ~9°/~8° 实证余量）。
REAL_INTERFERE_J4_MAX = 100.0
REAL_INTERFERE_J5_MIN = 165.0
# ★★★ v15.2（2026-11-03）：【J4 单独硬禁区 |J4|>150】
#   背景：v15 把 J4 限位 150→178 之后，P5 的规划解从 J4=123.60° 变成 J4=172.88°（11-03 11:14:37 实录），
#         ⇒ 实机报「断连收尾后未到位…173.19…误差0.84°」，界面显示姿态自干涉 ✗（= 用户说的"原本没有的自干涉"）
#   现有组合禁区 (|J4|>100 且 |J5|>165) 抓不住它：P5 的 J5 只有 58.81° ⇒ 不在禁区 ⇒ 放行 ⇒ 踩雷 ✗
#   ⇒ 新增：|J4| > 150 一律视为禁区（与 v14w23 的"实证安全族 |J4|≤95、150 留 55° 余量"一致）
#   ⇒ 效果：J4 限位仍是 178（能出解、不误杀"没有限位内的逆解"），但【选中的解 J4 必 ≤150】
#          ⇒ P5 回到 J4=123.60 的原解 ⇒ 既出解又不自干涉 ✓
REAL_INTERFERE_J4_HARD = 150.0


def _real_interfere_combo(q):
    """v14w26：关节是否落入实机自干涉组合禁区（J4×J5 耦合，控制器 -40006）。
    v15.2：追加 |J4|>150 的单独硬禁区（治 P5 的 J4=172.88 自干涉）。"""
    if abs(q[3]) > REAL_INTERFERE_J4_HARD:
        return True
    return abs(q[3]) > REAL_INTERFERE_J4_MAX and abs(q[4]) > REAL_INTERFERE_J5_MIN


def _real_limit_ok(q, lower, upper):
    """v14w22：关节目标是否同时满足模型限位与实机限位。"""
    for j in range(min(6, len(q))):
        lo = max(float(lower[j]), -REAL_JOINT_LIMITS[j])
        hi = min(float(upper[j]), REAL_JOINT_LIMITS[j])
        if not lo <= float(q[j]) <= hi:
            return False
    return True


def _try_set_tool_user():
    """Unsupported through this driver: RunCodeCustom becomes RunScript, not raw Tool/User."""
    raise ControllerMotionFault('当前驱动未验证Tool/User透传；禁止通过项目调用设置坐标系。')


def _movl_digit_safe_joints(q_target):
    """v14w：直发位姿数字净化 —— 控制器 MovL 参数校验 -30001 防御。

    实证（控制器 logs/all/log）：
      11:38:20 拒收 MovL(-0.000000,…,300.000000,90.000000,0.000000,-0.000000)
               → [MovL#820] the type of params is wrong: -30001
      15:55:51 接受 MovL(0.000000,…,299.999986,89.999995,-0.000003,0.000000) → return 0
    触发器（同目标、不同关节末位 ⇒ 不同参数形态 ⇒ 校验翻转）：
      x 负零/极小负 · rx 恰=+90.000000 · **三角(rx/ry/rz)负零——ry=-0 是 -30005 实锤**
      （10-15 09:16 与 10-14 拒收样本共同点；接受样本 ry 均为 +0）· rz=+180（保留防御）
      —— 同时设防，且只在零/边界区动手：
      · x ∈ (-0.01, 0.001) mm → 推到 ≥ +0.001（FK 位置与欧拉约定无关，可靠）
      · rx ∈ [89.999, 90.001] → 拉出该区（Pose_2_Fanuc 的 rx 与两份实录一致）
      · rz 为负零 (-0.0) → 推离
    手法：对发送关节贪心微扰（步长 0.0005°→0.05°，单关节累计 ≤0.05°，末端位移 ≲0.6mm
    ≪ 圆柱真裕度 19.9mm ≪ 法兰验收 8mm）；到位/法兰验收/MoveJ 收口仍对【原始认证关节】
    判定，收口回认证构型 —— 几何语义不变。P5 类非边界参数零扰动（首查即过，原样返回）。
    返回 (send_q, note)：无违规=(原关节,None)；成功=(微扰关节,说明)；失败=(None,原因)。"""
    def _digits(q):
        # v14w19：先按驱动下发格式（6位小数）定型再判——控制器校验的是字符串形态；
        # 客户端 Fanuc 与驱动在零点附近的正负号约定不一致，故三角一律推离零域。
        # v14w24：净化微扰可能把限位边界关节（如 J6=-360.00）推出模型限位，
        # SolveFK 会抛 TargetReachError——捕获后返回 None=不可行候选（评分置顶永不选中）。
        try:
            return [float('%.6f' % v) for v in Pose_2_Fanuc(robot.SolveFK(q))]
        except Exception:
            return None

    def _score(vals):
        if vals is None:
            return 1e9   # 越界候选：永不优于当前
        x, rx, ry, rz = vals[0], vals[3], vals[4], vals[5]
        s = 0.0
        if -0.01 < x < 0.001:                      # 零附近（含 -0.000000）且未达 +0.001
            s += (0.001 - x) / 0.001
        if 89.999 <= rx <= 90.001:                 # 恰卡 +90 边界（含 90.000000 整）
            s += (rx - 89.999) / 0.001
        # v14w19：三角必须整体离开零域 ≥0.001°——"-0.000000"形态是 -30005 实锤
        #（10-15 09:16/09:35 两次实录 ry 打印 -0.000000 均拒；-2e-7 打印即 -0.000000
        #  而浮点 !=0.0 会漏判；推离零域后客户端/驱动符号一致为正）
        for v in (rx, ry, rz):
            if abs(v) < 0.001:
                s += 1.0 + (0.001 - abs(v)) / 0.001
        if rz >= 179.999:                          # rz=+180 疑似越界（保留防御）
            s += 1.0 + (rz - 179.999) / 0.001
        return s

    base = list(q_target)
    cur = _score(_digits(base))
    if cur <= 0.0:
        return q_target, None
    q = list(base)
    solved = False
    for step in (0.0005, 0.002, 0.01, 0.05):
        improved = True
        while cur > 0.0 and improved:
            improved = False
            for j in range(6):
                for sgn in (1.0, -1.0):
                    q2 = q[:]
                    q2[j] += sgn * step
                    if abs(q2[j] - base[j]) > 0.05 + 1e-9:
                        continue
                    sc = _score(_digits(q2))
                    if sc < cur - 1e-12:
                        q, cur, improved = q2, sc, True
                        break
                if improved:
                    break
        if cur <= 0.0:
            solved = True
            break
    if not solved:
        return None, '发送位姿净化失败（边界参数 x/rx/rz 微调不出安全区）'
    touched = ['%s%+.4f' % ('J%d' % (k + 1), q[k] - base[k]) for k in range(6)
               if abs(q[k] - base[k]) > 1e-9]
    return q, '发送关节微扰 %s°（Δmax 对应末端 ≪1mm）：规避 -30001 边界参数；验收/收口仍回认证构型' \
        % ' '.join(touched)


def _movl_flange_accept(joints_now, joints_target):
    """v14q：直发 MovL 落点的法兰位姿级粗验收。

    v14p 首航实证：控制器 MovL 固有落点残差 ~5mm/0.6° 级（v14p 4.61mm/0.616°、v14l 5.5mm，
    双样本跨版本一致）——关节级 0.5° 判据会把正常落点误判为事故。改用法兰语义验收：
    FK(实测) vs FK(目标)，位置≤MOVL_FLANGE_TOL_MM 且姿态≤MOVL_FLANGE_TOL_DEG 即过；
    过后在 _execute_checked_real 里发一条 MoveJ 微纠偏收口（关节级 0.5° 校验罩住终点）。
    超容差=落点异常（构型翻转/卡住/送错目标），照旧抛 RuntimeError 即停待判读。"""
    _f_now = invH(robot.PoseFrame()) * robot.SolveFK(joints_now)      # 法兰位姿（无工具）
    _f_tgt = invH(robot.PoseFrame()) * robot.SolveFK(joints_target)
    _d = _f_now * invH(_f_tgt)
    _mm = norm(_d.Pos())
    _deg = math.degrees(pose_angle(_d))
    return _mm, _deg


def _movl_direct_ready():
    """v14p 法兰补偿MOVL 开关是否可用：GUI 变量已建（正常运行）才开；
    离线 verify 的 exec 命名空间里没有 real_movldirect_var（NameError），
    自动回 False——离线验证的计划/指纹与该开关无关（规划层零改动）。"""
    try:
        return isinstance(real_movldirect_var, tk.BooleanVar)
    except Exception:
        return False


MOVE_SEGMENT_MAX_DEG = 64.0  # 每瓣最大关节跨度：驱动约8秒无完成回报即断连，20°/s下64°≈3秒，留足裕量


J6_SPIN_SEGMENT_DEG = 60.0   # MoveL 纯J6自转段分瓣跨度（无平移时关节插值=笛卡尔路径）


def _is_pure_j6_spin(start, target):
    """MoveL 目标仅 J6 变化（J1~J5 不动）：关节插值与笛卡尔路径重合，可精确分瓣。"""
    return max(abs(a - b) for a, b in zip(start[:5], target[:5])) < 1e-6


def _move_with_completion_check(method, target, allow_split=True):
    """长运动分瓣执行（v9）：驱动对单条指令约8秒无完成回报就断连（本环境常态，
    test.py 同款假报，它每段部在几秒内完成所以从没撞上）；大跨度关节运动沿
    预检验证过的同一条关节直线剖成若干瓣，每瓣都在死线内完成，路径不变，
    仅增设停顿点。MoveL 纯J6自转段同理分瓣；带平移 MoveL 与小跨度段保持原样。"""
    if not allow_split:
        # v11: 单点运动/关节运动不分瓣，恢复一指令直达（到位校验与假断连容忍保留）
        _single_move_settle(method, target)
        return
    try:
        start = _live_joints()
        total = max(abs(float(b) - float(a)) for a, b in zip(start, target))
    except Exception:
        start, total = None, None
    if method == 'MoveJ' and total is not None and total > MOVE_SEGMENT_MAX_DEG:
        pieces = int(math.ceil(total / MOVE_SEGMENT_MAX_DEG))
        log('长运动分瓣：跨度%.1f° → %d 瓣执行（同一关节直线，仅增设停顿点）。' % (total, pieces))
        for k in range(1, pieces + 1):
            way = [a + (b - a) * k / pieces for a, b in zip(start, target)]
            _single_move_settle('MoveJ', way)
            _require_joints(way)  # 瓣间校验到位，也给驱动链路留出响应时间
        return
    if (method == 'MoveL' and total is not None and _is_pure_j6_spin(start, target)
            and total > J6_SPIN_SEGMENT_DEG):
        pieces = int(math.ceil(total / J6_SPIN_SEGMENT_DEG))
        log('J6自转分段：跨度%.1f° → %d 段MoveL（纯自转，路径与笛卡尔路径重合）。' % (total, pieces))
        for k in range(1, pieces + 1):
            way = [a + (b - a) * k / pieces for a, b in zip(start, target)]
            _single_move_settle('MoveL', way)
            _require_joints(way)
        return
    _single_move_settle(method, target)


_real_running = False  # 2026-10-09 补回：旧版 L510 有此初始化，升级版漏带导致点击即 NameError 静默炸裂


def _ensure_canonical_tool():
    """v14w17：工具坐标守护——检测到 identity(0)（存档僵尸/直发残留）自动恢复规范值并大声记日志。
    实发两次：2026-10-14 18:2x、2026-10-15 09:0x（归零→种子/P2 预检异常、P5 直发异常）。
    v14w39：同时恢复被直发窗口残留隐藏的门把手（GUI 中途被杀会留下隐藏态→预检漏检）。
    每次执行入口 + 程序启动各调一次；非零值不干预（可能正在被人工调整）。"""
    if _tool_window_depth:
        return False  # Do not undo the intentional identity TCP during MOVL.
    pose = robot.PoseTool()
    fixed = False
    canonical = Fanuc_2_Pose(list(CANONICAL_TOOL))
    if _same_tool_pose(pose, eye(4)) or _same_tool_pose(pose, canonical):
        tcp = _named_tool(TCP_TOOL_NAME, canonical)
        _restore_tool(canonical, tcp)
    if _same_tool_pose(pose, eye(4)):
        log('⚠️ 工具坐标为0（存档残留/直发残留）——已自动恢复 [0,0,130]，请确认后再跑。')
        fixed = True
    try:
        _gh = RDK.Item('门把手_bs1')
        if _gh.Valid() and not _gh.Visible():
            _gh.setVisible(True)
            log('⚠️ 门把手网格处于隐藏态（直发窗口残留）——已恢复显示。')
            fixed = True
    except Exception:
        pass
    return fixed


def _execute_checked_real(data, single_method=None):
    global _real_running
    log('【入口】_execute_checked_real：%d 点，single_method=%s' % (len(data) if data is not None else -1, single_method))
    if _real_running:
        log('已有实机任务正在执行。')
        return
    _real_running = True
    completed = 0
    movl_direct = False  # v14p：入口预置，防异常早于赋值时 except 块二次 NameError（v14l 教训）
    try:
        _ensure_canonical_tool()  # Failure must pass through task cleanup.
        log('开始校验录入数据…')
        records = _validated_records(data)
        log('录入数据校验通过：%d 点。' % len(records))
        if single_method is None and len(records) > 1:
            expanded = _retreat_orientation_records(records)
            log('连续轨迹：%d个录入点展开为%d个执行点（含姿态退让）。' % (len(records), len(expanded)))
            records = expanded
        deviation = float(real_deviation_var.get())
        if not math.isfinite(deviation) or deviation < 0:
            raise ValueError('允许偏离必须为非负有限数。')
        log('偏离上限 %.1f mm，检查机器人连接…' % deviation)
        if not ensure_connected():
            return
        start = _live_joints()
        log('实机当前关节：%s' % ['%.2f' % v for v in start])
        # 长预检/运动期间 RoboDK 主程序忙或不消费驱动输出，驱动链路会饿死断开（15:20:56 P1 中途断连同因）。
        # 保活线程用独立 API 连接（避免被 MoveJ 阻塞主连接），每2秒一次 ConnectedState（只读），
        # 贯穿预检+执行全程，直到任务结束才停（v7 错在预检后就停，P1 运动中饿死驱动）。
        import threading as _th
        _keepalive_stop = _th.Event()
        def _driver_keepalive():
            n = 0
            _ka_rdk = Robolink()
            _ka_robot = _ka_rdk.Item(robot.Name(), ITEM_TYPE_ROBOT)
            while not _keepalive_stop.wait(2.0):
                n += 1
                try:
                    s, _m = _ka_robot.ConnectedState()
                    if s < 0:
                        log('【保活】第%d次发现驱动掉线（%s），已请求重连。' % (n, _m))
                        _ka_robot.Connect()
                except Exception:
                    pass  # 主程序忙时 API 调用可能慢/超时，下一轮再试
        _ka_thread = _th.Thread(target=_driver_keepalive, daemon=True, name='driver_keepalive')
        _ka_thread.start()
        log('已启驱动保活（贯穿预检+执行）。')
        frame, tool = robot.PoseFrame(), robot.PoseTool()
        log('开始台子/地面避障预检，尚未发送运动指令。')
        plan = _prepare_real_plan(records, start, deviation, single_method)
        # 保活线程不在此处停：执行阶段同样需要（v7 教训）
        # 预检后复核：驱动必须就绪且关节与预检起始一致，否则取消。
        if not ensure_connected():
            log('预检后驱动断连，重连未成功，取消执行。')
            return
        _require_joints(start)
        log('预检后连接复核通过，准备发运动指令。')
        # v14w22：实机限位最后防线（规划器已过滤，此处兜底拦截任何漏网目标）
        # ★ v15（2026-11-03）：判限位前先做【同角归一化】—— 修一次误拦：
        #   实录 11:07:59 `段6 目标关节超出实机限位：['64.99','77.69','-96.48','198.78','64.99','0.00']`
        #   而 198.78° 与 −161.22° 是【同一个角】（差 360°），规划期用的是 −161.22（合法 ✓），
        #   最后防线却拿 198.78 去比 ⇒ 误判超限 ⇒ 整段 0 点即停 ✗。
        #   ⇒ 对每个关节先试 ±360k 的等价表示，取限位内的那个；都不在限位内才判死。
        #   ⇒ 并把归一化后的值【写回 plan】，避免执行时把 198.78 发给控制器（J6 合法域 ±360，故按轴各自限位判）。
        _lo, _hi, _ = robot.JointLimits()
        _lo, _hi = _lo.list(), _hi.list()

        def _nearest_in_limit(q):
            out = []
            for j in range(6):
                v = float(q[j])
                lo = max(float(_lo[j]), -REAL_JOINT_LIMITS[j])
                hi = min(float(_hi[j]), REAL_JOINT_LIMITS[j])
                if lo <= v <= hi:
                    out.append(v)
                    continue
                picked = None
                for k in (-1.0, 1.0):
                    alt = v + 360.0 * k
                    if lo <= alt <= hi:
                        picked = alt
                        break
                out.append(picked if picked is not None else v)
            return out

